// TwinCAT 3 PLC project WFServer
// ProgramVersion: 3.1.4026.14
// libraries:
//   Tc2_Standard, * (Beckhoff Automation GmbH)
//   Tc2_System, * (Beckhoff Automation GmbH)
//   Tc2_TcpIp, * (Beckhoff Automation GmbH)
//   Tc2_Utilities, * (Beckhoff Automation GmbH)
//   Tc3_Acsi, * (Beckhoff Automation GmbH)
//   Tc3_Ber, * (Beckhoff Automation GmbH)
//   Tc3_Collections, * (Beckhoff Automation GmbH)
//   Tc3_EventLogger, * (Beckhoff Automation GmbH)
//   Tc3_Gse, * (Beckhoff Automation GmbH)
//   Tc3_iec61850, * (Beckhoff Automation GmbH)
//   Tc3_iec61850_8_1, * (Beckhoff Automation GmbH)
//   Tc3_Mms, * (Beckhoff Automation GmbH)
//   Tc3_Rfc1006, * (Beckhoff Automation GmbH)
//   Tc3_Sockets, * (Beckhoff Automation GmbH)
//   Tc3_Tpkt, * (Beckhoff Automation GmbH)
//   Tc3_Ulosi, * (Beckhoff Automation GmbH)
// project tree:
//   / CommHandlerTask.TcTTO, DH_TCP_TX_TASK.TcTTO, IEC61850_TASK.TcTTO, UDP_RX_TASK.TcTTO, UDP_TX_TASK.TcTTO
//   DUTs/IEC61850/ E_DirectControlState.TcDUT, E_SboControlState.TcDUT
//   DUTs/IEC61850/User61850Enums/ E_ClrOp.TcDUT, E_CtlMd.TcDUT, E_TurCtl.TcDUT
//   DUTs/ S_TURBINECMD.TcDUT, S_TURBINEDATA.TcDUT
//   DUTs/TCP_UDP/ E_TCPConnectionState.TcDUT, E_UDPClientServerState.TcDUT, ST_TCPBinaryFrame.TcDUT, ST_TCPBinaryHeader.TcDUT, ST_UDPFrameEntry.TcDUT, TCP_DATA.TcDUT, UDP_DATA.TcDUT
//   GVLs/ CONSTANTS.TcGVL, TCP_GLOBALS.TcGVL, TcTelecontrol.TcGVL, UDP_GLOBALS.TcGVL
//   POUs/Common/ FB_LogFifo.TcPOU
//   POUs/COMM/ F_CreateTurbineCMD.TcPOU, F_InsertTurbineDataIEC61850.TcPOU, ParseTurbineData.TcPOU
//   POUs/ DH_TX_TCP_MAIN.TcPOU, P_IEC61850_MAIN.TcPOU, P_COMM_HANDLER.TcPOU, UDP_RX_MAIN.TcPOU, UDP_TX_MAIN.TcPOU
//   POUs/IEC61850Server/ FB_Control.TcPOU, FB_DirectControl.TcPOU, FB_DirectControlEnhanced.TcPOU, FB_SboControl.TcPOU, FB_SboControlEnhanced.TcPOU, FB_WTURBINEGse.TcPOU, FB_WTURBINEServerSession.TcPOU, FB_IEC61850.TcPOU, F_IEC61850ServerInit.TcPOU
//   POUs/IEC61850Server/User61850Enums/ FB_ClrOp.TcPOU, FB_CtlMd.TcPOU, FB_TurCtl.TcPOU
//   POUs/IEC61850Server/Util/ F_BuildAPTitle.TcPOU, F_BuildSelector.TcPOU, F_UdintToStringPadded.TcPOU
//   POUs/IEC61850Server/WTURBINE/ FB_IED_WTURBINE.TcPOU
//   POUs/IEC61850Server/WTURBINE/LD0/ FB_LD_WTURBINELD0.TcPOU
//   POUs/IEC61850Server/WTURBINE/LD0/LLN0/CDCs/ FB_DO_WTURBINE_LD0_LLN0_Beh.TcPOU, FB_DO_WTURBINE_LD0_LLN0_Health.TcPOU, FB_DO_WTURBINE_LD0_LLN0_Mod.TcPOU, FB_DO_WTURBINE_LD0_LLN0_NamPlt.TcPOU
//   POUs/IEC61850Server/WTURBINE/LD0/LLN0/ FB_LN_WTURBINE_LD0_LLN0.TcPOU
//   POUs/IEC61850Server/WTURBINE/LD0/LPHD1/CDCs/ FB_DO_WTURBINE_LD0_LPHD1_PhyHealth.TcPOU, FB_DO_WTURBINE_LD0_LPHD1_PhyNam.TcPOU, FB_DO_WTURBINE_LD0_LPHD1_Proxy.TcPOU
//   POUs/IEC61850Server/WTURBINE/LD0/LPHD1/ FB_LN_WTURBINE_LD0_LPHD1.TcPOU
//   POUs/IEC61850Server/WTURBINE/LD0/WALM1/CDCs/ FB_DO_WTURBINE_LD0_WALM1_Beh.TcPOU
//   POUs/IEC61850Server/WTURBINE/LD0/WALM1/ FB_LN_WTURBINE_LD0_WALM1.TcPOU
//   POUs/IEC61850Server/WTURBINE/LD0/WCNV1/CDCs/ FB_DO_WTURBINE_LD0_WCNV1_Beh.TcPOU, FB_DO_WTURBINE_LD0_WCNV1_Torq.TcPOU
//   POUs/IEC61850Server/WTURBINE/LD0/WCNV1/ FB_LN_WTURBINE_LD0_WCNV1.TcPOU
//   POUs/IEC61850Server/WTURBINE/LD0/WGEN1/CDCs/ FB_DO_WTURBINE_LD0_WGEN1_Beh.TcPOU, FB_DO_WTURBINE_LD0_WGEN1_RotSpd.TcPOU
//   POUs/IEC61850Server/WTURBINE/LD0/WGEN1/ FB_LN_WTURBINE_LD0_WGEN1.TcPOU
//   POUs/IEC61850Server/WTURBINE/LD0/WMET1/CDCs/ FB_DO_WTURBINE_LD0_WMET1_Beh.TcPOU, FB_DO_WTURBINE_LD0_WMET1_HorWdDir.TcPOU, FB_DO_WTURBINE_LD0_WMET1_HorWdSpd.TcPOU
//   POUs/IEC61850Server/WTURBINE/LD0/WMET1/ FB_LN_WTURBINE_LD0_WMET1.TcPOU
//   POUs/IEC61850Server/WTURBINE/LD0/WPPD1/CDCs/ FB_DO_WTURBINE_LD0_WPPD1_Beh.TcPOU, FB_DO_WTURBINE_LD0_WPPD1_ClrOp.TcPOU, FB_DO_WTURBINE_LD0_WPPD1_ClrOp_st.TcPOU, FB_DO_WTURBINE_LD0_WPPD1_DevOp.TcPOU, FB_DO_WTURBINE_LD0_WPPD1_DevOp_st.TcPOU, FB_DO_WTURBINE_LD0_WPPD1_DevSt.TcPOU, FB_DO_WTURBINE_LD0_WPPD1_DevSt_st.TcPOU
//   POUs/IEC61850Server/WTURBINE/LD0/WPPD1/DataSets/ FB_DS_TEMPLATE_LD1_WPPD1_ds01.TcPOU
//   POUs/IEC61850Server/WTURBINE/LD0/WPPD1/ FB_LN_WTURBINE_LD0_WPPD1.TcPOU
//   POUs/IEC61850Server/WTURBINE/LD0/WROT1/CDCs/ FB_DO_WTURBINE_LD0_WROT1_Beh.TcPOU, FB_DO_WTURBINE_LD0_WROT1_BlPthAngTgt.TcPOU, FB_DO_WTURBINE_LD0_WROT1_BlPthAngVal.TcPOU, FB_DO_WTURBINE_LD0_WROT1_RotSpd.TcPOU
//   POUs/IEC61850Server/WTURBINE/LD0/WROT1/ FB_LN_WTURBINE_LD0_WROT1.TcPOU
//   POUs/IEC61850Server/WTURBINE/LD0/WTUR1/CDCs/ FB_DO_WTURBINE_LD0_WTUR1_Beh.TcPOU, FB_DO_WTURBINE_LD0_WTUR1_DmdWSpt.TcPOU, FB_DO_WTURBINE_LD0_WTUR1_DmdWSpt_val.TcPOU, FB_DO_WTURBINE_LD0_WTUR1_TotWh.TcPOU, FB_DO_WTURBINE_LD0_WTUR1_TotWh_cntVal.TcPOU, FB_DO_WTURBINE_LD0_WTUR1_TurCtl.TcPOU, FB_DO_WTURBINE_LD0_WTUR1_TurCtl_st.TcPOU, FB_DO_WTURBINE_LD0_WTUR1_TurOp.TcPOU, FB_DO_WTURBINE_LD0_WTUR1_TurOp_st.TcPOU, FB_DO_WTURBINE_LD0_WTUR1_TurSt.TcPOU, FB_DO_WTURBINE_LD0_WTUR1_TurSt_st.TcPOU, FB_DO_WTURBINE_LD0_WTUR1_W.TcPOU
//   POUs/IEC61850Server/WTURBINE/LD0/WTUR1/ FB_LN_WTURBINE_LD0_WTUR1.TcPOU
//   POUs/IEC61850Server/WTURBINE/LD0/WYAW1/CDCs/ FB_DO_WTURBINE_LD0_WYAW1_Beh.TcPOU, FB_DO_WTURBINE_LD0_WYAW1_CabWup.TcPOU, FB_DO_WTURBINE_LD0_WYAW1_YwAng.TcPOU, FB_DO_WTURBINE_LD0_WYAW1_YwAngSpt.TcPOU, FB_DO_WTURBINE_LD0_WYAW1_YwAngSpt_val.TcPOU
//   POUs/IEC61850Server/WTURBINE/LD0/WYAW1/ FB_LN_WTURBINE_LD0_WYAW1.TcPOU
//   POUs/TCP/ FB_TCPClientConnection.TcPOU, FB_TCPClient.TcPOU, FB_TCPClientApplication.TcPOU
//   POUs/TCP/Util/ FB_TCPFrameFifo.TcPOU
//   POUs/UDP/ FB_UDPRxStateMachine.TcPOU, FB_UDPTxStateMachine.TcPOU
//   POUs/UDP/Util/ FB_UDPFrameFIFO.TcPOU
// real-time tasks:
//   TASK UDP_RX_TASK: cycle T#10ms, priority 15, ADS port 351
//   TASK CommHandlerTask: cycle T#10ms, priority 18, ADS port 353
//   TASK UDP_TX_TASK: cycle T#10ms, priority 2, ADS port 352
//   TASK IEC61850_TASK: cycle T#10ms, priority 1, ADS port 350
//   TASK DH_TCP_TX_TASK: cycle T#10ms, priority 3, ADS port 354
// I/O:
//   DEVICE GSE (RT-Ethernet Adapter) (disabled)

CONFIGURATION WFServer
    RESOURCE PLC ON TwinCAT3
        TASK CommHandlerTask(INTERVAL := T#10ms, PRIORITY := 18);
        TASK DH_TCP_TX_TASK(INTERVAL := T#10ms, PRIORITY := 3);
        TASK IEC61850_TASK(INTERVAL := T#10ms, PRIORITY := 1);
        TASK UDP_RX_TASK(INTERVAL := T#10ms, PRIORITY := 15);
        TASK UDP_TX_TASK(INTERVAL := T#10ms, PRIORITY := 2);
        PROGRAM P_COMM_HANDLER WITH CommHandlerTask : P_COMM_HANDLER;
        PROGRAM DH_TX_TCP_MAIN WITH DH_TCP_TX_TASK : DH_TX_TCP_MAIN;
        PROGRAM P_IEC61850_MAIN WITH IEC61850_TASK : P_IEC61850_MAIN;
        PROGRAM UDP_RX_MAIN WITH UDP_RX_TASK : UDP_RX_MAIN;
        PROGRAM UDP_TX_MAIN WITH UDP_TX_TASK : UDP_TX_MAIN;
    END_RESOURCE
END_CONFIGURATION

// ---- DUTs/IEC61850/E_DirectControlState.TcDUT
{attribute 'qualified_only'}
{attribute 'strict'}
TYPE E_DirectControlState : 
(
	Ready := 0,
	WaitForActivationTime := 1,
	PerformTest := 2,
	WaitForExecution := 3,
	Operate := 4,
	WaitForChange := 5,
	MirrorBlockedCommand := 6
) ;
END_TYPE

// ---- DUTs/IEC61850/E_SboControlState.TcDUT
{attribute 'qualified_only'}
{attribute 'strict'}
TYPE E_SboControlState : 
(
	Unselected := 0,
	Select_PerformTest := 1,
	WaitForSelection := 2,
	Ready := 3,
	WaitForActivationTime := 4,
	PerformTest := 5,
	WaitForExecution := 6,
	MirrorBlockedCommand := 7,
	Operate := 8,
	WaitForChange := 9,
	EndSelection := 10
) ;
END_TYPE

// ---- DUTs/IEC61850/User61850Enums/E_ClrOp.TcDUT
{attribute 'qualified_only'}
{attribute 'strict'}
TYPE E_ClrOp : 
(
	e_0 := 0, (*None*)
	e_1 := 1 (*Clear*)
) SINT;
END_TYPE

// ---- DUTs/IEC61850/User61850Enums/E_CtlMd.TcDUT
{attribute 'qualified_only'}
{attribute 'strict'}
TYPE E_CtlMd : 
(
	e_1 := 1, (*local*)
	e_2 := 2, (*remote*)
	e_3 := 3, (*auto*)
	e_4 := 4 (*test*)
) SINT;
END_TYPE

// ---- DUTs/IEC61850/User61850Enums/E_TurCtl.TcDUT
{attribute 'qualified_only'}
{attribute 'strict'}
TYPE E_TurCtl : 
(
	e_1 := 1, (*ROSCO*)
	e_2 := 2 (*Lio*)
) SINT;
END_TYPE

// ---- DUTs/S_TURBINECMD.TcDUT
(* Holds the command for all turbines *)
{attribute 'pack_mode' := '1'}
TYPE S_TURBINECMD :
STRUCT
	bEnable 		: ARRAY[1..c_nNumTurbines] OF BOOL;
	bEmergencyStop	: ARRAY[1..c_nNumTurbines] OF BOOL;
	eCtrlMode		: ARRAY[1..c_nNumTurbines] OF SINT;		// 1 Byte
	fWSpt			: ARRAY[1..c_nNumTurbines] OF REAL;
	fYawSpt			: ARRAY[1..c_nNumTurbines] OF REAL;
END_STRUCT
END_TYPE

// ---- DUTs/S_TURBINEDATA.TcDUT
{attribute 'pack_mode' := '1'}
TYPE S_TURBINEDATA :
STRUCT
	WindSpeed			: REAL;
	WindDirection		: REAL;
	PowerGen			: REAL;
	YawAng				: REAL;
	RotorSpeed			: REAL;
	PitchAngle			: REAL;
	PitchAngleSpt		: REAL;
	GenTorque			: REAL;
END_STRUCT
END_TYPE

// ---- DUTs/TCP_UDP/E_TCPConnectionState.TcDUT
TYPE E_TCPConnectionState :
(
	eTCP_STATE_IDLE,
	eTCP_STATE_CONNECT_START,
	eTCP_STATE_CONNECT_WAIT,
	eTCP_STATE_DATAEXCHANGE,
	eTCP_STATE_CLOSE_START,
	eTCP_STATE_CLOSE_WAIT,
	eTCP_STATE_ERROR
);
END_TYPE

// ---- DUTs/TCP_UDP/E_UDPClientServerState.TcDUT
TYPE E_UDPClientServerState :
(
	eUDP_STATE_IDLE		:= 0,
	eUDP_STATE_CREATE_START,
	eUDP_STATE_CREATE_WAIT,
	eUDP_STATE_SEND_START,
	eUDP_STATE_SEND_WAIT,
	eUDP_STATE_RECEIVE_START,
	eUDP_STATE_RECEIVE_WAIT,
	eUDP_STATE_CLOSE_START,
	eUDP_STATE_CLOSE_WAIT,
	eUDP_STATE_ERROR
);
END_TYPE

// ---- DUTs/TCP_UDP/ST_TCPBinaryFrame.TcDUT
(* Simple binary TCP/IP frame (8 byte aligned) *)
TYPE ST_TCPBinaryFrame :
STRUCT
	head	: ST_TCPBinaryHeader;(* Frame header (16 byte) *)
	data 	: TCP_DATA;(* User data (?? byte) *)

	(* Total frame size = 16+?? byte *)
END_STRUCT
END_TYPE

// ---- DUTs/TCP_UDP/ST_TCPBinaryHeader.TcDUT
(* Simple binary TCP/IP frame header (8 byte aligned) *)
TYPE ST_TCPBinaryHeader :
STRUCT
	dwStart		: DWORD	:= 16#BECF1234;	(* Start bytes *)
	cbLength	: UDINT(0..cTCP_BUFFER_SIZE) := 0;(* Max. length of attached binary data *)
	nS			: UDINT := 0;(* Send counter *)
	nR			: UDINT	:= 0;(* Receive counter *)
	
	(* Total header data size = 16 byte *)
END_STRUCT
END_TYPE

// ---- DUTs/TCP_UDP/ST_UDPFrameEntry.TcDUT
TYPE ST_UDPFrameEntry :
STRUCT
	stRemoteAddr 	: ST_SockAddr;	(* Remote address. String containing an (Ipv4) Internet Protocol dotted address and port number. *)
	sMessage		: UDP_DATA;	(* UDP packet data *)
END_STRUCT
END_TYPE

// ---- DUTs/TCP_UDP/TCP_DATA.TcDUT
// TYPE TCP_DATA : ARRAY[1..cTCP_FrameSize] OF BYTE; END_TYPE
TYPE TCP_DATA :
STRUCT
	nID				: UDINT;
	nUnixTime		: ULINT;
	YwAng			: REAL;
	YwAngSpt		: REAL;
	W				: REAL;
	WSpt			: REAL;
	HorWdSpd		: REAL;
	HorWdDir		: REAL;
	RotSpd			: REAL;
	PitchAngle		: REAL;
	PitchAngleSpt	: REAL;
// 	GenTorque		: REAL;
END_STRUCT
END_TYPE

// ---- DUTs/TCP_UDP/UDP_DATA.TcDUT
TYPE UDP_DATA : ARRAY[1..SIZEOF(S_TURBINECMD)*c_nNumTurbines] OF BYTE; END_TYPE

// ---- GVLs/CONSTANTS.TcGVL
VAR_GLOBAL CONSTANT
	c_nNumTurbines	: UDINT := 9;
	
	(* IEC 61850 Server Definitions *)
	c_aIpAddr 		: STRING := '172.19.3.190';
	c_aMMSPortBase 	: UDINT := 102;
	c_aAP_invIDBase : INT := 0;
	c_nNumSessions	: UINT := 1;
	
	(* UDP Connection Constants *)
	sSrvNetId			: T_AmsNetID 	:= '';(* TwinCAT TCP/IP server network address. Default: empty string. *)
	sLocalHost			: T_IPv4Addr 	:= '172.19.3.190';(* Local address: String containing an (Ipv4) Internet Protocol dotted address. *)
	nLocalTxPort		: UDINT			:= 11000;	(* UDP port used for transmission *)
	nLocalRxPort		: UDINT			:= 11001;	(* UDP port used for receiving *)
	sRemoteHost			: T_IPv4Addr 	:= '172.19.3.43';(* Remote address: String containing an (Ipv4) Internet Protocol dotted address. *)
	nRemoteTxPort		: UDINT 		:= 11000; (* Remote address: IP Tx port number. *)
	nRemoteRxPort		: UDINT			:= 10000; (* Remote address: IP Rx port number. *)
	
	UDP_RX_BUFFER_SIZE 	: UDINT := c_nNumTurbines * 1024; 	// Size of the UDP RX FIFO Buffer in Bytes
	UDP_TX_BUFFER_SIZE 	: UDINT := 1024; 	// Size of the UDP TX FIFO Buffer in Bytes
	
	UDP_ERR_TX_FIFO_OF	: UDINT := 16#8103;
	UDP_ERR_RX_FIFO_OF	: UDINT := 16#8104;
END_VAR

// ---- GVLs/TCP_GLOBALS.TcGVL
VAR_GLOBAL CONSTANT
	cTCP_BUFFER_SIZE						: UDINT := 1000;
	cTCP_FrameSize							: UDINT := 256;

	cTCP_SEND_CYCLE_TIME					: TIME := T#1S;
	cTCP_RECEIVE_POLLING_TIME		 		: TIME := T#100MS;
	cTCP_RECEIVE_TIMEOUT					: TIME := T#50S;

	(* Some project specific error codes *)
	cTCP_ERROR_RECEIVE_TIMEOUT				: UDINT := 16#8101;(* Receive timeout error *)
	cTCP_ERROR_SENDFIFO_OVERFLOW			: UDINT := 16#8102;(* Send fifo overflow *)
	cTCP_ERROR_RECFIFO_OVERFLOW				: UDINT := 16#8103;(* Receive fifo overflow *)
	cTCP_ERROR_INVALID_FRAME_FORMAT		: UDINT := 16#8104;(* Invalid frame format/data *)
END_VAR

// ---- GVLs/TcTelecontrol.TcGVL
VAR_GLOBAL
	ipCreator: I_AcsiCodeCreatorClass := GVL_AcsiVars.Creator.SetCodeRev(codeRev:=7).SetGuiVer(major:=3, minor:=98, build:=20, revision:=0);
	
	(* IEC61850 Data Models for Turbine *)
	fbWTURBINE: ARRAY[1..c_nNumTurbines] OF FB_IED_WTURBINE;
	
	(* IEC61850 Server Objects, one for each turbine *)
	fbServer : ARRAY[1..c_nNumTurbines] OF FB_iec61850ServerClass;
	
	(* IEC61850 Server Sessions, one or multiple for each server object *)
	fbSession: ARRAY[1..c_nNumTurbines, 1..c_nNumSessions] OF FB_WTURBINEServerSession;
	
// 	{warning 'Please configure your server IP-address in the initialization code of the server function block below:'}
	(* Server container *)
// 	fbWTURBINEServer: FB_iec61850ServerClass := (ipIED:=fbWTURBINE, settings:=(bEnable:=TRUE, sLocalHost:='192.168.1.100', nCalled_AP_InvID:=0, nCalling_AP_InvID:=0, nCalled_AE_InvID:=0, nCalling_AE_InvID:=0));
	
	(* Server connections *)
// 	fbWTURBINEServerSession1: FB_WTURBINEServerSession := (fbConnection:=(ipServer:=fbWTURBINEServer, settings:=(bEnable:=TRUE)));
	(*
	fbWTURBINEServerSession2: FB_WTURBINEServerSession := (fbConnection:=(ipServer:=fbWTURBINEServer, settings:=(bEnable:=TRUE)));
	...
	fbWTURBINEServerSessionN: FB_WTURBINEServerSession := (fbConnection:=(ipServer:=fbWTURBINEServer, settings:=(bEnable:=TRUE)));
	*)
	
	
// 	fbWTURBINEGse: FB_WTURBINEGse := (fbAdapter:=(ipIED:=fbWTURBINE, settings:=(sMulticastAddr:='01-0C-CD-01-00-00', eDispatchMode:=E_GseDispatchMode.NonPromiscuous)));
	
	
END_VAR

// ---- GVLs/UDP_GLOBALS.TcGVL
VAR_GLOBAL
	(* Global TX and RX buffers, together with their respective critical section handlers*)
// 	fbUDP_RX_CS			: FB_IecCriticalSection;
	fbRxFIFO			: FB_UDPFrameFIFO;
	
// 	fbUDP_TX_CS			: FB_IecCriticalSection;
	fbTxFIFO			: FB_UDPFrameFIFO;
END_VAR

// ---- POUs/P_COMM_HANDLER.TcPOU
PROGRAM P_COMM_HANDLER
VAR
	i					: UDINT;
	nAddr				: ULINT;
	stReceivedFrom		: ST_UDPFrameEntry;
	sLoggedMessage		: UDP_DATA;
	dVal_1				: LREAL;
	dVal_2				: LREAL;	
	sTurbineData		: S_TURBINEDATA;
	iTemp				: ULINT;
	
	sTxTimer			: TON;
	bSend				: BOOL := FALSE;
	cTxTimerPeriod		: TIME := T#500MS;
	sTurbineCmd			: S_TURBINECMD;
	stSendTo			: ST_UDPFrameEntry;;
END_VAR


(* First we pop from the UDP RX buffer, and process the received data accordingly *)
REPEAT
	fbRxFIFO.RemoveHead( );
	IF fbRxFIFO.bOk THEN

		(* TODO:: Implement received frame handler *)
		stReceivedFrom := fbRxFIFO.stGet;
		IF stReceivedFrom.stRemoteAddr.sAddr = sRemoteHost AND stReceivedFrom.stRemoteAddr.nPort = nRemoteTxPort THEN
// 			sLoggedMessage := stReceivedFrom.sMessage;
			nAddr := 0;
			FOR i := 1 TO c_nNumTurbines DO
				sTurbineData := ParseTurbineData(ADR(stReceivedFrom.sMessage) + nAddr);
				F_InsertTurbineDataIEC61850(nID := i, sTurbineData := sTurbineData);
				nAddr := nAddr + SIZEOF(S_TURBINEDATA);
			END_FOR
		END_IF
// 		MEMCPY(ADR(dVal_1), ADR(sLoggedMessage), SIZEOF(dVal_1));
// 		MEMCPY(ADR(dVal_2), ADR(sLoggedMessage) + SIZEOF(dVal_1), SIZEOF(dVal_2));
// 			ADSLOGSTR( ADSLOG_MSGTYPE_HINT OR ADSLOG_MSGTYPE_LOG OR ADSLOG_MSGTYPE_MSGBOX, '%s', stReceivedFrom.sMessage );
		
	END_IF
UNTIL NOT fbRxFIFO.bOk
END_REPEAT


(* Second, we take the turbine setpoints and transmit to the turbine *)
bSend := sTxTimer.Q;
sTxTimer(IN := NOT sTxTimer.Q, PT := cTxTimerPeriod);

IF bSend THEN
	sTurbineCmd := F_CreateTurbineCMD();
	fbTXFIFO.AddTail( );
	iTemp :=  SIZEOF(sTurbineCmd);
	MEMCPY(ADR(stSendTo.sMessage), ADR(sTurbineCmd), SIZEOF(sTurbineCmd));
	stSendTo.stRemoteAddr.sAddr := sRemoteHost;	(* Remote host IP address *)
	stSendTo.stRemoteAddr.nPort := nRemoteRxPort;	(* Remote host port number *)
	fbTxFIFO.AddTail( stPut := stSendTo );
END_IF

END_PROGRAM

// ---- POUs/COMM/ParseTurbineData.TcPOU
FUNCTION ParseTurbineData
VAR_INPUT
	sMessage		: POINTER TO BYTE;
END_VAR
VAR_OUTPUT
	sTurbineData	: S_TURBINEDATA;
// 	bOk				: BOOL;
END_VAR
VAR
	i				: UDINT;
	nAddr			: ULINT;
END_VAR

// bOk := FALSE;
MEMCPY(ADR(sTurbineData), sMessage, SIZEOF(sTurbineData));
// nAddr := 0;
// MEMCPY(ADR(sTurbineData.WindSpeed) + nAddr, sMessage + nAddr, SIZEOF(sTurbineData.WindSpeed));
// nAddr := nAddr + SIZEOF(sTurbineData.WindSpeed);
// 
// MEMCPY(ADR(sTurbineData.WindDirection), sMessage + nAddr, SIZEOF(sTurbineData.WindDirection));
// nAddr := nAddr + SIZEOF(sTurbineData.WindDirection);
// 
// MEMCPY(ADR(sTurbineData.PowerGen), sMessage + nAddr, SIZEOF(sTurbineData.PowerGen));
// nAddr := nAddr + SIZEOF(sTurbineData.PowerGen);
// 
// MEMCPY(ADR(sTurbineData.YawAng), sMessage + nAddr, SIZEOF(sTurbineData.YawAng));
// nAddr := nAddr + SIZEOF(sTurbineData.YawAng);
// 
// MEMCPY(ADR(sTurbineData.RotorSpeed), sMessage + nAddr, SIZEOF(sTurbineData.RotorSpeed));
// nAddr := nAddr + SIZEOF(sTurbineData.RotorSpeed);
// 
// MEMCPY(ADR(sTurbineData.PitchAngle), sMessage + nAddr, SIZEOF(sTurbineData.PitchAngle));
// nAddr := nAddr + SIZEOF(sTurbineData.PitchAngle);
// 
// MEMCPY(ADR(sTurbineData.PitchAngleSpt), sMessage + nAddr, SIZEOF(sTurbineData.PitchAngleSpt));
// nAddr := nAddr + SIZEOF(sTurbineData.PitchAngleSpt);
// 
// MEMCPY(ADR(sTurbineData.GenTorque), sMessage + nAddr, SIZEOF(sTurbineData.GenTorque));
// nAddr := nAddr + SIZEOF(sTurbineData.GenTorque);

// bOk := TRUE;

END_FUNCTION

// ---- POUs/COMM/F_InsertTurbineDataIEC61850.TcPOU
FUNCTION F_InsertTurbineDataIEC61850
VAR_INPUT
	nID				: UDINT;
	sTurbineData	: S_TURBINEDATA;
END_VAR
VAR_OUTPUT
END_VAR
VAR
END_VAR

IF nID >= 1 OR nID <= c_nNumTurbines THEN
	fbWTURBINE[nID].WTURBINELD0.WMET1.HorWdSpd.mag.fValue := sTurbineData.WindSpeed;
	fbWTURBINE[nID].WTURBINELD0.WMET1.HorWdDir.mag.fValue := sTurbineData.WindDirection;
	fbWTURBINE[nID].WTURBINELD0.WTUR1.W.mag.fValue := sTurbineData.PowerGen;
	fbWTURBINE[nID].WTURBINELD0.WYAW1.YwAng.mag.fValue := sTurbineData.YawAng;
	fbWTURBINE[nID].WTURBINELD0.WROT1.RotSpd.mag.fValue := sTurbineData.RotorSpeed;
	fbWTURBINE[nID].WTURBINELD0.WROT1.BlPthAngVal.mag.fValue := sTurbineData.PitchAngle;
	fbWTURBINE[nID].WTURBINELD0.WROT1.BlPthAngTgt.mag.fValue := sTurbineData.PitchAngleSpt;
 	fbWTURBINE[nID].WTURBINELD0.WCNV1.Torq.mag.fValue := sTurbineData.GenTorque;
END_IF

END_FUNCTION

// ---- POUs/COMM/F_CreateTurbineCMD.TcPOU
FUNCTION F_CreateTurbineCMD
VAR_INPUT
// 	nID				: UDINT;
END_VAR
VAR_OUTPUT
	sTurbineCmd		: S_TURBINECMD;
END_VAR
VAR
	temp: SINT;
	nID: UDINT;
END_VAR


FOR nID := 1 TO c_nNumTurbines DO
	temp := fbWTURBINE[nID].WTURBINELD0.WTUR1.TurOp.st_.stVal.iAny;
	sTurbineCmd.bEnable[nID] :=  SINT_TO_BOOL(temp);
	sTurbineCmd.bEmergencyStop[nID] := FALSE;
	sTurbineCmd.eCtrlMode[nID] := fbWTURBINE[nID].WTURBINELD0.WTUR1.TurCtl.st_.stVal.iAny;
	sTurbineCmd.fWSpt[nID] 	:= fbWTURBINE[nID].WTURBINELD0.WTUR1.DmdWSpt.val.mxVal.fValue;
	sTurbineCmd.fYawSpt[nID] := fbWTURBINE[nID].WTURBINELD0.WYAW1.YwAngSpt.val.mxVal.fValue;
END_FOR

END_FUNCTION

// ---- POUs/DH_TX_TCP_MAIN.TcPOU
PROGRAM DH_TX_TCP_MAIN
VAR
	sSrvNetID 	: T_AmsNetID := '';(* TwinCAT TCP/IP server network address *)
	bEnable 	: BOOL := TRUE;(* TRUE => Enable client data exchange, FALSE => Disable *)	
	
	bLog		: BOOL := TRUE;(* TRUE => Enable message/error log, FALSE => Disable*)
	
	fbClient : FB_TCPClient := ( sRemoteHost:= '172.19.3.214',(* IP address of remote server! *)
								nRemotePort:= 9003,(* Port number of remote server! *)
								sPrefix := 'CLIENT1::' );(* TCP/IP client (connection) instance *)
								
	fbCloseAll		: FB_SocketCloseAll;
	bInitialize		: BOOL := TRUE;
END_VAR

IF fbCloseAll.bBusy OR fbCloseAll.bError THEN
	RETURN;
END_IF
bInitialize := FALSE;

fbClient( sSrvNetID := sSrvNetID, bEnable := bEnable, bLog := bLog );

END_PROGRAM

// ---- POUs/TCP/FB_TCPClient.TcPOU
FUNCTION_BLOCK FB_TCPClient
VAR_INPUT
	sSrvNetID	: T_AmsNetID	:= '';(* TwinCAT TCP/IP server network address *)
	sRemoteHost	: T_IPv4Addr 	:= '127.0.0.1';(* Server IP network address *)
	nRemotePort	: UDINT 		:= 200;(* Server port number *)
	bEnable		: BOOL 			:= FALSE;(* TRUE => enable client data exchange, FALSE => disable *)
	bLog		: BOOL 			:= FALSE;(* TRUE => Enable log message output, FALSE => Disable *)
	sPrefix		: STRING 		:= 'CLIENT::';(* Log message description string (allows the identification of log message source) *)
END_VAR
VAR_OUTPUT
	eState		: E_SocketConnectionState := eSOCKET_DISCONNECTED;(* TCP/IP connection state *)
END_VAR
VAR
	fbApplication 	: FB_TCPClientApplication;(* Client application control function block *)
	fbConnection	: FB_TCPClientConnection;(* Client data exchange control function block *)
	fbTx 			: FB_TCPFrameFifo;(* Tx fifo *)
	fbRx 			: FB_TCPFrameFifo;(* Rx fifo *)
	fbLog			: FB_LogFifo;(* Log/debug/error fifo *)
END_VAR

(*-------------------------- Trigger data exchange -----------------------------------------------*)
fbConnection( 	sSrvNetID := sSrvNetID, fbRx := fbRx, fbTx := fbTx, fbLog := fbLog, 
				bEnable := bEnable, sRemoteHost := sRemoteHost, nRemotePort := nRemotePort,  
				bLog := bLog, sPrefix := sPrefix, eState=>eState );
	
IF fbConnection.eState = eSOCKET_CONNECTED THEN(* Connection established *)
	fbApplication( fbTx := fbTx, fbRx := fbRx, fbLog := fbLog );
END_IF

END_FUNCTION_BLOCK

// ---- POUs/TCP/FB_TCPClientApplication.TcPOU
FUNCTION_BLOCK FB_TCPClientApplication
VAR_IN_OUT
	fbTx 		: FB_TCPFrameFifo;(* TX fifo *)
	fbRx 		: FB_TCPFrameFifo;(* RX fifo *)
	fbLog		: FB_LogFifo;(* Log message fifo *)
END_VAR
VAR
	stToServer	: TCP_DATA;
	stFromServer: TCP_DATA;
	sLogMessage	: T_MaxString := '';
	nCounter	: UDINT;
	fbSndTimer	: TON;
	i: UDINT;
	fbFormat   : FB_FormatString;
	sFormatted : T_MaxString;
	
	
	fbTime   : FB_LocalSystemTime := ( bEnable := TRUE, dwCycle := 1 );
	sTime 	: T_MaxString;
 	nDataLen     : INT;
    nUnixTime    : LINT;
END_VAR

(*------------------- Send cyclic message strings ------------------------------------*)
(* TODO: Make this 'application/task' agnostic. *)
(* For now, it always sends logging data to the historian *)
fbSndTimer( IN := TRUE, PT := cTCP_SEND_CYCLE_TIME );
IF fbSndTimer.Q THEN(* Send string to server *)
	fbSndTimer( IN := FALSE );

// 	nCounter := nCounter  + 1;
// 	stToServer := MAXSTRING_TO_BYTEARR(CONCAT( 'Client message: ', UDINT_TO_STRING(nCounter) ));
//  
// 	fbTx.AddTail( stPut := stToServer );(* Put string to the tx fifo *)
// 	IF NOT fbTx.bOk THEN(* TX fifo overflow => log error *)
// 		fbLog.Error( sMessage := 'FB_FrameFifo(sender)\0', nErrID := cTCP_ERROR_SENDFIFO_OVERFLOW );
// 	END_IF
	
	fbTime();
	sTime := SYSTEMTIME_TO_STRING(fbTime.systemTime);
	FOR i := 1 TO c_nNumTurbines DO
		
		stToServer.nID := i;
		stToServer.nUnixTime := (F_GetSystemTime() - 116444736000000000) / 10000000;
		stToServer.YwAng := fbWTURBINE[i].WTURBINELD0.WYAW1.YwAng.mag.fValue;
		stToServer.YwAngSpt := fbWTURBINE[i].WTURBINELD0.WYAW1.YwAngSpt.val.mxVal.fValue;
		stToServer.W := fbWTURBINE[i].WTURBINELD0.WTUR1.W.mag.fValue;
		stToServer.WSpt := fbWTURBINE[i].WTURBINELD0.WTUR1.DmdWSpt.val.mxVal.fValue;
		stToServer.HorWdSpd := fbWTURBINE[i].WTURBINELD0.WMET1.HorWdSpd.mag.fValue;
		stToServer.HorWdDir := fbWTURBINE[i].WTURBINELD0.WMET1.HorWdDir.mag.fValue;
		stToServer.RotSpd := fbWTURBINE[i].WTURBINELD0.WROT1.RotSpd.mag.fValue;
		stToServer.PitchAngle := fbWTURBINE[i].WTURBINELD0.WROT1.BlPthAngVal.mag.fValue;
		stToServer.PitchAngleSpt := fbWTURBINE[i].WTURBINELD0.WROT1.BlPthAngTgt.mag.fValue;
// 		stToServer.GenTorque := fbWTURBINE[i].WTURBINELD0.WROT1.
		
		
		
		
		fbTx.AddTail( stPut := stToServer );(* Put string to the tx fifo *)
		IF NOT fbTx.bOk THEN(* TX fifo overflow => log error *)
			fbLog.Error( sMessage := 'FB_FrameFifo(sender)\0', nErrID := cTCP_ERROR_SENDFIFO_OVERFLOW );
		END_IF
	END_FOR

END_IF

END_FUNCTION_BLOCK

// ---- POUs/TCP/Util/FB_TCPFrameFifo.TcPOU
(* Tx/Rx (string data) fifo control function block *)
FUNCTION_BLOCK FB_TCPFrameFifo
VAR_INPUT
	bLog		: BOOL		:= FALSE;(* TRUE => Enable log message output, FALSE => Disable *)
	sPrefix		: STRING	:= 'Unknown::';(* Log message description string (allows the identification of log message source) *)
	stPut		: TCP_DATA;(* Frame to add (write) to the fifo *)
END_VAR
VAR_OUTPUT
	bOk			: BOOL; 	(* TRUE = New entry added or removed succesfully, FALSE = Fifo overflow or fifo empty *)
	stGet		: TCP_DATA;(* Frame removed (read) from fifo *)
	nCount		: UDINT		:= 0;(* Number of fifo entries *)
	cbFree		: UDINT 	:= 0;(* Free buffer space *)
END_VAR
VAR
	fbBuffer 	: FB_MemRingBuffer;(* Basic (lower level) buffer control function block *)
	buffer		: ARRAY[-3..cTCP_BUFFER_SIZE] OF BYTE;(* Internal buffer memory *)
END_VAR

;

ACTION AddTail:
(* Adds new fifo entry *)
fbBuffer.A_AddTail( pBuffer:= ADR(buffer), cbBuffer:= SIZEOF(buffer),
					pWrite := ADR( stPut ), cbWrite := SIZEOF( stPut ), 
					bOk=>bOk, nCount=>nCount );
IF bOk THEN
	cbFree := cTCP_BUFFER_SIZE - fbBuffer.cbSize;(* Calculate the free buffer space *)
// 	IF bLog THEN(* Log message *)
// 		F_ADSLOGHEXDATA( CONCAT( sPrefix, '<=' ), ADR( stPut ), SIZEOF( stPut ) );
// 	END_IF
END_IF
END_ACTION

ACTION Clear:
(* Resets fifo = clears all data *)
MEMSET( ADR( stGet ), 0, SIZEOF( stGet ) );
fbBuffer.A_Reset( pBuffer:= ADR(buffer), cbBuffer:= SIZEOF(buffer),
					pWrite := ADR( stPut ), cbWrite := SIZEOF( stPut ), 
					pRead := ADR( stGet ), cbRead := SIZEOF( stPut ),
					bOk=>bOk, nCount=>nCount );
cbFree := cTCP_BUFFER_SIZE;(* Free buffer size *)
END_ACTION

ACTION RemoveHead:
(* Removes oldest fifo entry *)
MEMSET( ADR( stGet ), 0, SIZEOF( stGet ) );
fbBuffer.A_RemoveHead( pBuffer:= ADR(buffer), cbBuffer:= SIZEOF(buffer),
						pRead := ADR( stGet ), cbRead := SIZEOF( stGet ),
						bOk=>bOk, nCount=>nCount );
IF bOk THEN
	cbFree := cTCP_BUFFER_SIZE - fbBuffer.cbSize;(* Calculate the free buffer space *)
END_IF
END_ACTION

END_FUNCTION_BLOCK

// ---- POUs/Common/FB_LogFifo.TcPOU
(* Log/debug/error message fifo *)
FUNCTION_BLOCK FB_LogFifo
VAR_INPUT
	bLog		: BOOL 		:= FALSE;(* TRUE => Enable log message output, FALSE => Disable *)
	sPrefix		: STRING 	:= 'Unknown::';(* Log message description string (allows the identification of log message source) *)
	
	sMessage	: STRING 	:= '';(* String message to add (write) to the fifo *)
	nErrID		: UDINT 	:= 0;(* Error code to add (write) to the fifo *)
	hSocket		: T_HSOCKET;(* Socket connection handle *)
END_VAR
VAR_OUTPUT
	bOk			: BOOL;(* TRUE = New entry added or removed succesfully, FALSE = Fifo overflow or fifo empty *)
	sGet		: T_MaxString := '';(* String entry removed (read) from fifo *)
	nCount		: UDINT := 0;(* Number of fifo entries *)
END_VAR
VAR
	fbBuffer 	: FB_StringRingBuffer;(* Basic (lower level) string buffer control function block *)
	buffer		: ARRAY[0..cTCP_BUFFER_SIZE] OF BYTE;(* Internal buffer memory *)
	sSource		: T_MaxString;	
	sPut		: T_MaxString;
END_VAR

;

ACTION Clear:
(* Clears all fifo entries *)
fbBuffer.A_Reset( 	pBuffer := ADR( buffer ), cbBuffer := SIZEOF( buffer ), 
					bOk=>bOk, nCount=>nCount, getValue=>sGet );
END_ACTION

ACTION Error:
(* Adds new fifo entry *)
IF nErrID = 0 THEN
	sSource := '::Error: 0x';
ELSIF ( nErrID AND 16#80000000) = 16#80000000 THEN
	IF nErrID = 16#80072746 THEN
		sSource := '::Win32 error (the connection is reset by remote side): 0x';
	ELSE
		sSource := '::Win32 error: 0x';
	END_IF
ELSIF (nErrID AND 16#00008100) = 16#00008100 THEN
	CASE nErrID OF
		cTCP_ERROR_RECEIVE_TIMEOUT:
			sSource := '::PLC sample project receive timeout error: 0x';
		cTCP_ERROR_SENDFIFO_OVERFLOW:
			sSource := '::PLC sample project send fifo overflow error: 0x';
		cTCP_ERROR_RECFIFO_OVERFLOW:
			sSource := '::PLC sample project receive fifo overflow error: 0x';
	ELSE
		sSource := '::Other PLC sample project error: 0x';
	END_CASE
ELSIF (nErrID AND 16#00008000) = 16#00008000 THEN
	sSource := '::Internal TCP/IP Connection Server error: 0x';
ELSE
	sSource := '::TwinCAT System error: 0x';
END_IF

sPut := CONCAT( CONCAT( CONCAT( sPrefix, sMessage ), sSource ), DWORD_TO_HEXSTR( nErrID AND 16#FFFF, 0, FALSE ) ); 

fbBuffer.A_AddTail( pBuffer:= ADR(buffer), cbBuffer:= SIZEOF(buffer),
					putValue:= sPut, bOk=>bOk, nCount=>nCount );
IF bOk THEN
	IF bLog THEN(* Log error message *)
		ADSLOGSTR( ADSLOG_MSGTYPE_ERROR OR ADSLOG_MSGTYPE_LOG, '%s', sPut );	
	END_IF
END_IF
END_ACTION

ACTION Message:
(* Adds new fifo entry *)
sPut := CONCAT( CONCAT( sPrefix, sMessage ), CONCAT( '::', HSOCKET_TO_STRING(hSocket) ) );
fbBuffer.A_AddTail( pBuffer:= ADR(buffer), cbBuffer:= SIZEOF(buffer),
					putValue:= sPut, bOk=>bOk, nCount=>nCount );
IF bOk THEN
	IF bLog THEN(* Log information message *)
		ADSLOGSTR( ADSLOG_MSGTYPE_HINT OR ADSLOG_MSGTYPE_LOG, '%s', sPut );	
	END_IF
END_IF
END_ACTION

ACTION Remove:
(* Removes oldest fifo entry *)
IF nCount = 0 THEN
	sGet := '';
	bOk := FALSE;
	RETURN;
END_IF

fbBuffer.A_RemoveHead( pBuffer:= ADR(buffer), cbBuffer:= SIZEOF(buffer),
						getValue=>sGet, bOk=>bOk, nCount=>nCount );
END_ACTION

END_FUNCTION_BLOCK

// ---- POUs/TCP/FB_TCPClientConnection.TcPOU
(* 	This function block implements simple TCP/IP client protocol. *)
FUNCTION_BLOCK FB_TCPClientConnection
VAR_IN_OUT
	fbTx 		: FB_TCPFrameFifo;(* TX fifo *)
	fbRx 		: FB_TCPFrameFifo;(* RX fifo *)
	fbLog		: FB_LogFifo;(* Log message fifo *)
END_VAR
VAR_INPUT
	sSrvNetID	: T_AmsNetID	:= '';(* TwinCAT TCP/IP server network address *)
	sRemoteHost	: T_IPv4Addr 	:= '127.0.0.1';(* IP address of remote server *)
	nRemotePort	: UDINT			:= 200;(* Remote server port *)
	bEnable		: BOOL			:= FALSE;(* TRUE => Enable/connect, FALSE => Disable/disconnect *)
	tReconnect	: TIME 			:= T#5S;(* Try to reconnect after this time *)
	bLog		: BOOL 			:= FALSE; (* TRUE => Enable debug output, FALSE => Disable debug output *)
	sPrefix		: STRING 		:= 'CLIENT::';(* Log message description string (allows the identification of log message source) *)
END_VAR
VAR_OUTPUT
	eState		: E_SocketConnectionState := eSOCKET_DISCONNECTED;(* TCP/IP connection state *)
END_VAR
VAR
	fbConnect 	: FB_ClientServerConnection;(* Create/release TCP/IP connection *)
	fbSend		: FB_SocketSend;(* Send TCP/IP data *)
	fbReceive	: FB_SocketReceive;(* Receive TCP/IP data *)
	nState 		: BYTE;(* Global state *)
	bSndBusy 	: BOOL;(* Tx state *)
	bRcvBusy 	: BOOL;(* Rx state *)
	bDisconnect	: BOOL;(* Disconnect flag, if set the socket will be closed *)

	fbPollTimer	: TON;(* Rx data poll timer *)
	fbResponseTimer	: TON;(* Response timeout timer *)
	fbReconnectTimer : TON;(* Reconnect timer *)

	nS			: UDINT;(* Send frame counter *)
	nR			: UDINT;(* Received frame counter *)
	cbReceived	: UDINT;(* Count of received data bytes *)
	rxBuffer	: ARRAY[0..cTCP_BUFFER_SIZE] OF BYTE;
	cbFrame		: UDINT;(* Rx frame byte size *)
	stTxFrame	: ST_TCPBinaryFrame;(* Tx frame buffer (inclusive header) *)
	stRxFrame	: ST_TCPBinaryFrame;(* Rx frame buffer (inclusive header) *)
	bAbort		: BOOL;(* Flag to abort frame parsing loop *)
	sSend: Tc2_System.T_MaxString;
END_VAR

CASE nState OF
	0:(* Create TCP/IP connection *)
		fbConnect( 	sSrvNetID 		:= sSrvNetID,
					nMode			:= SEL( bLog, 0, CONNECT_MODE_ENABLEDBG ),(* Enable/disable debug output *)
					sRemoteHost 	:= sRemoteHost,
					nRemotePort 	:= nRemotePort,
					tReconnect		:= tReconnect,
					bEnable			:= bEnable,
					eState			=> eState );
		IF NOT fbConnect.bBusy THEN
			IF NOT fbConnect.bError THEN
				IF eState = eSOCKET_CONNECTED THEN(* we are connected *)
					
					fbTx.Clear( sPrefix := CONCAT( sPrefix, 'FB_FrameFifo(sender)::' ), bLog := bLog );(* Clear TX fifo (optional) *)
					fbRx.Clear( sPrefix := CONCAT( sPrefix, 'FB_FrameFifo(receiver)::' ), bLog := bLog );(* Clear RX fifo (optional) *)
					fbLog.Clear( sPrefix := sPrefix, bLog := bLog );(* Clear log fifo (optional) *)
					bSndBusy := FALSE;
					bRcvBusy := FALSE;
					bDisconnect := FALSE;
					cbReceived 	:= 0;(* Reset number of received data bytes *)
					nR 			:= 0;(* Reset receive frame counter *)
					nS 			:= 0;(* Reset send frame counter *)

					fbPollTimer( IN := FALSE, PT := T#0S );
					fbResponseTimer( IN := FALSE, PT := cTCP_RECEIVE_TIMEOUT );
					fbReconnectTimer( IN := FALSE, PT := tReconnect );
				
					fbLog.Message( sMessage := 'Connection established!', hSocket := fbConnect.hSocket );
					nState 	:= 1;
				END_IF
			ELSE(* Connect error => log error *)
				fbLog.Error( sMessage := 'FB_ClientServerConnection()', nErrID := fbConnect.nErrId );
			END_IF
		END_IF


	1:(* Data exchange state *)
		bDisconnect := NOT bEnable OR bDisconnect;(* User/internal disconnect requested? *)
		IF bDisconnect AND NOT bSndBusy AND NOT bRcvBusy THEN
			bDisconnect := FALSE;
			fbLog.Message( sMessage := 'Closing connection!', hSocket := fbConnect.hSocket );
			nState := 2;(* Disconnect *)
		ELSE

			(* --------------------------- Send tx data --------------------------------- *)
			IF NOT bDisconnect AND NOT bSndBusy THEN
				fbTx.RemoveHead();(* Remove oldest user data entry *)
				IF fbTx.bOk THEN(* Success *)
						
					stTxFrame.data := fbTx.stGet;
					
					(* Append/create some protocol header *)
					stTxFrame.head.dwStart 	:= 16#BECF1234;(* Frame start bytes *)
					stTxFrame.head.cbLength := SIZEOF( stTxFrame.data);(* Set length of user data *)
					stTxFrame.head.nS 		:= nS;(* Number of send frames *)
					stTxFrame.head.nR 		:= nR;(* Number of received frames *)
					
					(* Send frame *)
					fbSend( bExecute := FALSE );
// 					sSend := BYTEARR_TO_MAXSTRING(stTxFrame.data);
					
					fbSend(	sSrvNetID 	:= sSrvNetID,
							hSocket		:= fbConnect.hSocket,
							cbLen		:= SIZEOF(TCP_DATA),(* Size of header + size of user data *)
							pSrc		:= ADR(stTxFrame.data),(* Pointer to the frame data *)
							bExecute	:= TRUE );
					bSndBusy := TRUE;
				END_IF
			ELSE(* Wait until send not busy *)
				fbSend( bExecute := FALSE );
				IF NOT fbSend.bBusy THEN
					bSndBusy := FALSE;
					IF NOT fbSend.bError THEN(* No error *)
						nS := nS + 1;(* Increment the number of send frames *)
					ELSE(* Send error => Log error and disconnect *)
						fbLog.Error( sMessage := 'FB_SocketSend()', nErrID := fbSend.nErrId );
						bDisconnect := TRUE;(* Set flag *)
					END_IF
				END_IF
			END_IF
			(* -------------------------------------------------------------------------- *)

// 			(* ------------------ Get/fetch rx data ------------------------------------- *)
// 			IF NOT bDisconnect AND NOT bRcvBusy THEN
// 				fbPollTimer( IN := TRUE );
// 				IF fbPollTimer.Q THEN
// 					IF fbRx.cbFree >= SIZEOF(stRxFrame.data) THEN(* Check free rx fifo space *)
// 						fbPollTimer( IN := FALSE, PT := cTCP_RECEIVE_POLLING_TIME );
// 						fbReceive( bExecute := FALSE );
// 						fbReceive( 	sSrvNetId	:= sSrvNetID,
// 									hSocket		:= fbConnect.hSocket,
// 									cbLen		:= SIZEOF(rxBuffer) - cbReceived,
// 									pDest		:= ADR(rxBuffer) + cbReceived,
// 									bExecute	:= TRUE );
// 						bRcvBusy := TRUE;
// 					END_IF
// 				END_IF
// 				
// 			ELSE(* Wait until receive not busy *)
// 				
// 				fbReceive( bExecute := FALSE );
// 				IF NOT fbReceive.bBusy THEN
// 					bRcvBusy := FALSE;
// 					IF NOT fbReceive.bError THEN
// 						IF fbReceive.nRecBytes > 0 THEN (* Some bytes received *)
// 
// 							fbPollTimer( IN := FALSE, PT := T#0S );(* Bytes received => increase the read (polling) speed *)
// 							fbResponseTimer( IN := FALSE );(* Bytes received => disable timeout check *)
// 							cbReceived := cbReceived + fbReceive.nRecBytes;
// 
// 							(* Parse received bytes *)
// 							REPEAT
// 								bAbort := TRUE;(* Set flag *)
// 								
// 								IF cbReceived >= SIZEOF(stRxFrame.head) THEN (* All header bytes received => check header data *)
// 									
// 									MEMCPY( ADR( stRxFrame.head ), ADR( rxBuffer ), SIZEOF( stRxFrame.head ) );(* Get header data *)
// 								
// 									IF (stRxFrame.head.dwStart = 16#BECF1234) (* Check start bytes *)
// 									AND (stRxFrame.head.nS = nR )(* Check counter (send counter == expected receive counter?) *)
// 									AND (stRxFrame.head.cbLength <= SIZEOF(stRxFrame.data))(* Check frame (user data) length *)
// 									THEN
// 									
// 										cbFrame := SIZEOF(stRxFrame.head) + stRxFrame.head.cbLength;(* Calculate the expected receive frame length *)
// 										IF cbReceived >= cbFrame  THEN (* All frame (user data) bytes received? *)
// 	
// 											MEMCPY( ADR( stRxFrame ), ADR( rxBuffer ), MIN( SIZEOF(stRxFrame), cbFrame ) );
// 											fbRx.AddTail( stPut := stRxFrame.data );(* Add user data to the rx fifo *)
// 											IF fbRx.bOk THEN
// 												nR := nR + 1;(* Increment receive counter *)
// 
// 												MEMMOVE( ADR( rxBuffer ), ADR( rxBuffer ) + cbFrame, cbReceived - cbFrame );(* Shift the remaining rx bytes *)
// 												cbReceived := cbReceived - cbFrame;(* Recalculate the size of the remaining rx bytes *)
// 
// 												IF fbRx.cbFree >= SIZEOF(stRxFrame.data) THEN
// 													bAbort := FALSE;(* reset flag, try to parse next frame *)
// 												END_IF
// 											ELSE (* Fifo overflow => log error and disconnect *)
// 												fbLog.Error( sMessage := 'FB_FrameFifo(receiver)', nErrID := cTCP_ERROR_RECFIFO_OVERFLOW );
// 												bDisconnect := TRUE;(* Set flag *)
// 												RETURN;
// 											END_IF
// 
// (*										ELSE repeat reading *)
// 										END_IF
// 
// 									ELSE(* Receive error => Invalid frame format/data *)
// 										fbLog.Error( sMessage := 'FB_ClientConnection()', nErrID := cTCP_ERROR_INVALID_FRAME_FORMAT );
// 										bDisconnect := TRUE;(* Set flag *)
// 										RETURN;
// 									END_IF
// 
// (*								ELSE repeat reading *)
// 								END_IF (* IF cbReceived >= SIZEOF(stRxFrame.head) THEN *)
// 
// 							UNTIL bAbort
// 							END_REPEAT
// 
// 						ELSE(* No bytes received *)
// 							fbResponseTimer( IN := TRUE );(* No bytes received => enable timeout check *)
// 							IF fbResponseTimer.Q THEN (* Timeout error*)
// 								fbResponseTimer( IN := FALSE );
// 								fbLog.Error( sMessage := 'FB_ClientConnection()', nErrID := cTCP_ERROR_RECEIVE_TIMEOUT );
// 								bDisconnect := TRUE;(* Set flag *)
// 							END_IF							
// 						END_IF(* IF fbReceive.nRecBytes > 0 THEN *)
// 
// 					ELSE(* Receive error => Log error and disconnect *)
// 						fbLog.Error( sMessage := 'FB_SocketReceive()', nErrID := fbReceive.nErrId );
// 						bDisconnect := TRUE;(* set flag *)
// 					END_IF
// 
// 				END_IF(* IF NOT fbReceive.bBusy THEN *)
// 				
// 			END_IF(* IF NOT bDisconnect AND NOT bRcvBusy THEN *)
// 			(* -------------------------------------------------------------------------- *)
			
			
		END_IF(* IF bDisconnect AND NOT bSndBusy AND NOT bRcvBusy THEN *)


	2:(* Disconnect *)
		fbConnect( bEnable:= FALSE, eState=>eState );
		IF eState = eSOCKET_DISCONNECTED THEN
			fbReconnectTimer( IN := TRUE );(* Please wait some seconds and then try to connect again *)
			IF fbReconnectTimer.Q THEN
				fbReconnectTimer( IN := FALSE );
				nState := 0;
			END_IF
		END_IF


END_CASE

END_FUNCTION_BLOCK

// ---- POUs/P_IEC61850_MAIN.TcPOU
PROGRAM P_IEC61850_MAIN
VAR
	fbIEC 	: FB_IEC61850;	
END_VAR

fbIEC();

END_PROGRAM

// ---- POUs/IEC61850Server/FB_IEC61850.TcPOU
FUNCTION_BLOCK FB_IEC61850
VAR
	bInitDone: BOOL := FALSE;	

	i: UDINT;
	j: UDINT;
END_VAR

IF NOT bInitDone THEN
	F_IEC61850ServerInit();

	bInitDone := TRUE;
END_IF

FOR i := 1 TO c_nNumTurbines DO
	fbServer[i].Execute();
	FOR j := 1 TO c_nNumSessions DO
		fbSession[i,j]();
	END_FOR
END_FOR

END_FUNCTION_BLOCK

// ---- POUs/IEC61850Server/F_IEC61850ServerInit.TcPOU
FUNCTION F_IEC61850ServerInit
VAR
	i: UDINT;
	j: UDINT;
END_VAR

FOR i := 1 TO c_nNumTurbines DO
	fbServer[i].ipIED := fbWTURBINE[i];
	
	
	fbServer[i].settings.bEnable := TRUE;
	fbServer[i].settings.sLocalHost := c_aIpAddr;
	fbServer[i].settings.nLocalPort := c_aMMSPortBase + i - 1;
	fbServer[i].settings.sCalled_T_Selector := F_BuildSelector(i);
	fbServer[i].settings.sCalled_S_Selector := F_BuildSelector(i);
	fbServer[i].settings.sCalled_P_Selector := CONCAT('00 00 ', F_UdintToStringPadded(i, 2));
	fbServer[i].settings.sCalled_AP_Title := F_BuildAPTitle(i);
	fbServer[i].settings.nCalled_AP_InvID := i;
	fbServer[i].settings.nCalled_AE_InvID := i;
	fbServer[i].settings.nCalling_AP_InvID := i - 1;
	fbServer[i].settings.nCalling_AE_InvID := i - 1;
	
	FOR j := 1 TO c_nNumSessions DO
		fbSession[i,j].fbConnection.ipServer := fbServer[i];
		fbSession[i,j].fbConnection.settings.bEnable := TRUE;
		fbSession[i,j].nID := i;
	END_FOR
	
	fbWTURBINE[i].WTURBINELD0.WPPD1.ds01.OnInit();
END_FOR

END_FUNCTION

// ---- POUs/IEC61850Server/Util/F_BuildSelector.TcPOU
FUNCTION F_BuildSelector : STRING
VAR_INPUT
    iValue : UDINT;
END_VAR

F_BuildSelector := CONCAT('00 ', F_UdintToStringPadded(iValue, 2));

END_FUNCTION

// ---- POUs/IEC61850Server/Util/F_UdintToStringPadded.TcPOU
FUNCTION F_UdintToStringPadded : STRING
VAR_INPUT
    iValue : UDINT;
    nWidth : DINT;
END_VAR

VAR
    sTemp : STRING(20);
END_VAR

sTemp := UDINT_TO_STRING(iValue);
WHILE LEN(sTemp) < nWidth DO
    sTemp := CONCAT('0', sTemp);
END_WHILE

F_UdintToStringPadded := sTemp;

END_FUNCTION

// ---- POUs/IEC61850Server/Util/F_BuildAPTitle.TcPOU
FUNCTION F_BuildAPTitle : STRING
VAR_INPUT
    iValue : UDINT;
END_VAR

F_BuildAPTitle := CONCAT('1.1.1.999.', UDINT_TO_STRING(iValue));

END_FUNCTION

// ---- POUs/UDP_RX_MAIN.TcPOU
PROGRAM UDP_RX_MAIN
VAR
	fbCloseAll 			: FB_SocketCloseAll;
   	bInitialize			: BOOL := TRUE;
	
	bEnable				: BOOL 			:= TRUE;(* TRUE => Enable/connect, FALSE => Disable/disconnect *)
	bLog				: BOOL			:= TRUE;(* TRUE => Enable log message output, FALSE => Disable *)
	
	fbRx				: FB_UDPRxStateMachine := (sPrefix := 'UDP_RX::');
END_VAR

(* On PLC reset or program download close all opened/created sockets *)
fbCloseAll( sSrvNetId := sSrvNetId, bExecute:= bInitialize );
IF fbCloseAll.bBusy OR fbCloseAll.bError THEN
	RETURN;
END_IF
// IF NOT fbCloseAll.nErrId THEN
//     RETURN; // Not done yet
// END_IF
bInitialize := FALSE;

fbRx(fbRxFifo:=fbRxFIFO, bEnable:=bEnable, bLog:=bLog);

END_PROGRAM

// ---- POUs/UDP/FB_UDPRxStateMachine.TcPOU
FUNCTION_BLOCK FB_UDPRxStateMachine
VAR_IN_OUT
	fbRxFIFO		: FB_UDPFrameFIFO;
END_VAR
VAR_INPUT
	bEnable			: BOOL			:= FALSE;
	tReconnect		: TIME			:= T#5S;
	bLog			: BOOL			:= FALSE;
	sPrefix			: STRING		:= 'UDP_RX::';
END_VAR
VAR_OUTPUT
	bCreated		: BOOL			:= FALSE;
END_VAR
VAR
	fbCreate		: FB_SocketUdpCreate;
	fbClose			: FB_SocketClose;
	hSocket			: T_HSOCKET;
	fbReceiveFrom	: FB_SocketUdpReceiveFrom;
	stReceivedFrom	: ST_UDPFrameEntry;
	fbCreateTimer	: TON := ( PT := T#0S );	
	eState			: E_UDPClientServerState;
END_VAR

CASE eState OF
	(* Idle State *)
	eUDP_STATE_IDLE:
		IF bEnable XOR bCreated THEN
			IF bEnable THEN
				(* Clear rx fifo *)
				fbRxFIFO.Clear( sPrefix := CONCAT( sPrefix, 'FB_FrameFifo(sender)::' ), bLog := bLog );
				
				(* At program start (first time) connect immediately, next time after delay time *)
				fbCreateTimer( IN := TRUE );
				IF fbCreateTimer.Q THEN
					fbCreateTimer( IN := FALSE, PT := tReconnect ); 
					eState := eUDP_STATE_CREATE_START;
				END_IF
			ELSE
				eState := eUDP_STATE_CLOSE_START;
			END_IF
		ELSIF bCreated THEN
			eState := eUDP_STATE_RECEIVE_START;
// 			fbRxFIFO.RemoveHead( stGet => stSendTo );
// 			IF fbRxFIFO.bOk THEN
// 				eState := eUDP_STATE_SEND_START;
// 			END_IF
		ELSE
			fbCreateTimer( IN := FALSE, PT := T#0S );
		END_IF
	
	(* Creation States *)
	eUDP_STATE_CREATE_START:
		fbCreate( bExecute := FALSE  );
		fbCreate( sSrvNetId := sSrvNetId, sLocalHost:= sLocalHost, nLocalPort:= nLocalRxPort, bExecute:= TRUE );
		eState := eUDP_STATE_CREATE_WAIT;

	eUDP_STATE_CREATE_WAIT:
		fbCreate( bExecute := FALSE );
		IF NOT fbCreate.bBusy THEN
			IF NOT fbCreate.bError THEN
				bCreated := TRUE;
				hSocket := fbCreate.hSocket;
// 				fbLog.Message( sMessage := 'Connectionless (UDP) socket created!', hSocket := fbCreate.hSocket );
				eState := eUDP_STATE_IDLE;
			ELSE
// 				fbLog.Error( sMessage := 'FB_SocketUdpCreate()', nErrID := fbCreate.nErrID );
				eState := eUDP_STATE_ERROR;
			END_IF
		END_IF
		
	eUDP_STATE_RECEIVE_START:
		MEMSET( ADR( stReceivedFrom ), 0, SIZEOF( stReceivedFrom ) );
		fbReceiveFrom( bExecute := FALSE );
		fbReceiveFrom( sSrvNetId := sSrvNetId, 
						pDest:= ADR( stReceivedFrom.sMessage ),
						cbLen:= SIZEOF( stReceivedFrom.sMessage ) - 1, (* Without string delimiter *)
						hSocket:= fbCreate.hSocket, bExecute:= TRUE );
		eState := eUDP_STATE_RECEIVE_WAIT;

	eUDP_STATE_RECEIVE_WAIT:
		fbReceiveFrom( bExecute := FALSE );
		IF NOT fbReceiveFrom.bBusy THEN
			IF NOT fbReceiveFrom.bError THEN
				IF fbReceiveFrom.nRecBytes > 0 THEN
					
					stReceivedFrom.stRemoteAddr.sAddr := fbReceiveFrom.sRemoteHost;
					stReceivedFrom.stRemoteAddr.nPort := fbReceiveFrom.nRemotePort;
					
					fbRxFIFO.AddTail( stPut := stReceivedFrom );
	// 				IF NOT fbRxFIFO.bOk THEN(* Check for fifo overflow *)
	// 					fbLog.Error( sMessage :='FB_FrameFifo(receiver)', nErrID := PLCPRJ_ERROR_RECFIFO_OVERFLOW );
	// 				END_IF
				END_IF
				eState := eUDP_STATE_IDLE;
			ELSE
	// 			fbLog.Error( sMessage := 'FB_SocketUdpReceiveFrom()', nErrID := fbReceiveFrom.nErrID );
				IF fbReceiveFrom.nErrID = 16#80072746 THEN(* Connection is reset by remote side *)
					eState := eUDP_STATE_IDLE;
				ELSE
					eState := eUDP_STATE_ERROR;
				END_IF
			END_IF
		END_IF
		
		
	(* Closing States *)
	eUDP_STATE_CLOSE_START:
// 		fbLog.Message( sMessage := 'Closing connectionless (UDP) socket!', hSocket := fbCreate.hSocket );
		fbClose( bExecute := FALSE );
		fbClose( sSrvNetId := sSrvNetId, hSocket := fbCreate.hSocket, bExecute := TRUE );
		eState := eUDP_STATE_CLOSE_WAIT;
		
	eUDP_STATE_CLOSE_WAIT:
		fbClose( bExecute := FALSE );
		IF NOT fbClose.bBusy THEN
			bCreated := FALSE;
			IF NOT fbClose.bError THEN
				eState := eUDP_STATE_IDLE;
			ELSE
// 				fbLog.Error( sMessage := 'FB_SocketClose()', nErrID := fbClose.nErrID );
				eState := eUDP_STATE_ERROR;
			END_IF
		END_IF

	(* Error State *)

	eUDP_STATE_ERROR: (* Error step *)
		IF bCreated THEN
			eState := eUDP_STATE_CLOSE_START;
		ELSE
			eState := eUDP_STATE_IDLE;
		END_IF
		
END_CASE

//FB_Exit must be implemented explicitly. If there is an implementation, then the
//method is called before the controller removes the code of the function block instance
//(implicit call). The return value is not evaluated.
METHOD FB_Exit: BOOL
VAR_INPUT
    bInCopyCode: BOOL;  // TRUE: the exit method is called in order to leave the instance which will be copied afterwards (online change).  
END_VAR
IF bCreated THEN
    fbClose(sSrvNetId := '', hSocket := hSocket, bExecute := TRUE);
END_IF
END_METHOD

END_FUNCTION_BLOCK

// ---- POUs/UDP/Util/FB_UDPFrameFIFO.TcPOU
(* Tx/Rx (string data) fifo control function block *)
FUNCTION_BLOCK FB_UDPFrameFIFO
VAR_INPUT
	bLog		: BOOL := FALSE;(* TRUE => Enable log message output, FALSE => Disable *)
	sPrefix		: STRING := 'Unknown::';(* Log message description string (allows the identification of log message source) *)
	stPut		: ST_UDPFrameEntry;(* Frame entry to add (write) to the buffer *)
END_VAR
VAR_OUTPUT
	bOk			: BOOL;(* TRUE = New entry added or removed succesfully, FALSE = Fifo overflow or fifo empty *)
	stGet		: ST_UDPFrameEntry;(* Frame entry removed (read) from fifo *)
	nCount		: UDINT := 0;(* Number of fifo entries *)
END_VAR
VAR
	fbBuffer 	: FB_MemRingBuffer;(* Basic (lower level) string buffer control function block *)
	buffer		: ARRAY[0..UDP_RX_BUFFER_SIZE] OF BYTE;(* Internal buffer memory *)
	fbCriticalSection:	FB_IecCriticalSection; (* Critical Section required for thread-safety *)
END_VAR

ACTION AddTail:
(* Adds new fifo entry *)
// IF fbCriticalSection.Enter() THEN
	fbBuffer.A_AddTail( pBuffer:= ADR(buffer), cbBuffer:= SIZEOF(buffer),
					pWrite:= ADR( stPut ), cbWrite := SIZEOF( stPut ), 
					bOk=>bOk, nCount=>nCount );
					
// 	fbCriticalSection.Leave();
// END_IF
// IF bOk AND bLog THEN(* Log message *)
// 	ADSLOGSTR( ADSLOG_MSGTYPE_HINT OR ADSLOG_MSGTYPE_LOG, 
// 			CONCAT( CONCAT( sPrefix, SOCKETADDR_TO_STRING(stPut.stRemoteAddr) ), '>>"%s"' ),
// 			stPut.sMessage );
// END_IF
END_ACTION

ACTION Clear:
(* Clears all fifo entries *)
// stGet.sMessage := 0;
// IF fbCriticalSection.Enter() THEN
	MEMSET(ADR(stGet.sMessage), 0, SIZEOF(stGet.sMessage));
	stGet.stRemoteAddr.nPort := 0;
	stGet.stRemoteAddr.sAddr := '';
	fbBuffer.A_Reset( pBuffer := ADR( buffer ), cbBuffer := SIZEOF( buffer ), bOk=>bOk, nCount=>nCount ); 
	
// 	fbCriticalSection.Leave();
// END_IF
END_ACTION

ACTION RemoveHead:
(* Removes oldest fifo entry *)

// IF fbCriticalSection.Enter() THEN
	IF nCount = 0 THEN
		MEMSET(ADR(stGet.sMessage), 0, SIZEOF(stGet.sMessage));
		stGet.stRemoteAddr.nPort := 0;
		stGet.stRemoteAddr.sAddr := '';
		bOk := FALSE;
		RETURN;
	END_IF
	
	fbBuffer.A_RemoveHead( pBuffer:= ADR(buffer), cbBuffer:= SIZEOF(buffer),
							pRead := ADR( stGet ), cbRead := SIZEOF( stGet ),
							bOk=>bOk, nCount=>nCount );
// 	fbCriticalSection.Leave();
// END_IF
END_ACTION

METHOD TEMPRemoveHead : BOOL
VAR_IN_OUT
	stGet	: ST_UDPFrameEntry;
END_VAR
VAR_INPUT
END_VAR
VAR_OUTPUT
	bOk		: BOOL;
END_VAR
IF fbCriticalSection.Enter() THEN
	IF nCount = 0 THEN
		MEMSET(ADR(stGet.sMessage), 0, SIZEOF(stGet.sMessage));
		stGet.stRemoteAddr.nPort := 0;
		stGet.stRemoteAddr.sAddr := '';
		bOk := FALSE;
		RETURN;
	END_IF
	
	fbBuffer.A_RemoveHead( pBuffer:= ADR(buffer), cbBuffer:= SIZEOF(buffer),
							pRead := ADR( stGet ), cbRead := SIZEOF( stGet ),
							bOk=>bOk, nCount=>nCount );
	fbCriticalSection.Leave();
END_IF
END_METHOD

END_FUNCTION_BLOCK

// ---- POUs/UDP_TX_MAIN.TcPOU
PROGRAM UDP_TX_MAIN
VAR
	bSendOnceToRemote	: BOOL;
	bEnable				: BOOL 			:= TRUE;(* TRUE => Enable/connect, FALSE => Disable/disconnect *)
	bLog				: BOOL			:= TRUE;(* TRUE => Enable log message output, FALSE => Disable *)
	
	fbTx				: FB_UDPTxStateMachine := (sPrefix := 'UDP_TX::');
	stSendTo			: ST_UDPFrameEntry;
	
	
	iTemp_1: BYTE := 1;
	iTemp_2: BYTE := 2;
	
	fbCloseAll 			: FB_SocketCloseAll;
	bInitialize: BOOL;
END_VAR

fbCloseAll( sSrvNetId := sSrvNetId, bExecute:= bInitialize );
IF fbCloseAll.bBusy OR fbCloseAll.bError THEN
	RETURN;
END_IF
bInitialize := FALSE;

fbTx(fbTxFifo:=fbTxFIFO, bEnable:=bEnable, bLog:=bLog);

// iTemp_1 := iTemp_1 + 1;
// iTemp_2 := iTemp_2+2;
// 
// IF fbTx.bCreated THEN
// 	IF bSendOnceToRemote THEN
// 		bSendOnceToRemote 			:= FALSE;		(* Clear flag *)
// 		MEMSET(ADR(stSendTo.sMessage), 0, SIZEOF(stSendto.sMessage));
// 		stSendTo.sMessage[1] := INT_TO_BYTE(iTemp_1);
// 		stSendTo.sMessage[2] := INT_TO_BYTE(iTemp_2);		
// 		stSendTo.stRemoteAddr.sAddr := sRemoteHost;	(* Remote host IP address *)
// 		stSendTo.stRemoteAddr.nPort := nRemoteTxPort;	(* Remote host port number *)
// 		fbTxFIFO.AddTail( stPut := stSendTo );	(* Add new entry to the send queue *)
// 	END_IF
// END_IF

END_PROGRAM

// ---- POUs/UDP/FB_UDPTxStateMachine.TcPOU
FUNCTION_BLOCK FB_UDPTxStateMachine
VAR_IN_OUT
	fbTxFIFO		: FB_UDPFrameFIFO;
END_VAR
VAR_INPUT
	bEnable			: BOOL			:= FALSE;			// TRUE => Enable/connect, FALSE => Disable/disconnect
	tReconnect		: TIME			:= T#5S;			// Reconnect delay time
	bLog			: BOOL			:= FALSE;			// TRUE => Enable log message output, FALSE => Disable 
	sPrefix			: STRING 		:= 'PeerToPeerX::'; // Log message description string (allows the identification of log message source)
END_VAR
VAR_OUTPUT
	bCreated		: BOOL;		// Connectionless socket state (TRUE => created, FALSE => closed)
END_VAR
VAR
	fbCreate		: FB_SocketUdpCreate;
	hSocket			: T_HSOCKET;
	fbClose			: FB_SocketClose;
	fbSendTo		: FB_SocketUdpSendTo;
	stSendTo		: ST_UDPFrameEntry;
	fbCreateTimer	: TON := ( PT := T#0S );	
	eState			: E_UDPClientServerState;
END_VAR

CASE eState OF
	(* Idle State *)
	eUDP_STATE_IDLE:
		IF bEnable XOR bCreated THEN
			IF bEnable THEN
				(* Clear send fifo *)
				fbTxFIFO.Clear( sPrefix := CONCAT( sPrefix, 'FB_FrameFifo(sender)::' ), bLog := bLog );
				
				(* At program start (first time) connect immediately, next time after delay time *)
				fbCreateTimer( IN := TRUE );
				IF fbCreateTimer.Q THEN
					fbCreateTimer( IN := FALSE, PT := tReconnect ); 
					eState := eUDP_STATE_CREATE_START;
				END_IF
			ELSE
				eState := eUDP_STATE_CLOSE_START;
			END_IF
		ELSIF bCreated THEN
			fbTxFIFO.RemoveHead( stGet => stSendTo );
			IF fbTxFIFO.bOk THEN
				eState := eUDP_STATE_SEND_START;
			END_IF
		ELSE
			fbCreateTimer( IN := FALSE, PT := T#0S );
		END_IF
	
	(* Creation States *)
	eUDP_STATE_CREATE_START:
		fbCreate( bExecute := FALSE  );
		fbCreate( sSrvNetId := sSrvNetId, sLocalHost:= sLocalHost, nLocalPort:= nLocalTxPort, bExecute:= TRUE );
		eState := eUDP_STATE_CREATE_WAIT;

	eUDP_STATE_CREATE_WAIT:
		fbCreate( bExecute := FALSE );
		IF NOT fbCreate.bBusy THEN
			IF NOT fbCreate.bError THEN
				bCreated := TRUE;
				hSocket := fbCreate.hSocket;
// 				fbLog.Message( sMessage := 'Connectionless (UDP) socket created!', hSocket := fbCreate.hSocket );
				eState := eUDP_STATE_IDLE;
			ELSE
// 				fbLog.Error( sMessage := 'FB_SocketUdpCreate()', nErrID := fbCreate.nErrID );
				eState := eUDP_STATE_ERROR;
			END_IF
		END_IF
	
	(* Sending States *)
	eUDP_STATE_SEND_START:
		fbSendTo( bExecute := FALSE );
		fbSendTo( sSrvNetId := sSrvNetId, sRemoteHost := stSendTo.stRemoteAddr.sAddr,
					nRemotePort := stSendTo.stRemoteAddr.nPort,
					pSrc:= ADR( stSendTo.sMessage ),
					//cbLen:= INT_TO_UDINT(LEN( stSendTo.sMessage )) + 1, (* Include the end delimiter *)
					cbLen := SIZEOF(UDP_DATA),
					hSocket:= fbCreate.hSocket, bExecute:= TRUE );
		eState := eUDP_STATE_SEND_WAIT;

	eUDP_STATE_SEND_WAIT:
		fbSendTo( bExecute := FALSE );
		IF NOT fbSendTo.bBusy THEN
			IF NOT fbSendTo.bError THEN
				eState := eUDP_STATE_IDLE;
			ELSE
// 				fbLog.Error( sMessage := 'FB_SocketUdpSendTo()', nErrID := fbSendTo.nErrID );
				eState := eUDP_STATE_ERROR;
			END_IF
		END_IF
		
	(* Closing States *)
	eUDP_STATE_CLOSE_START:
// 		fbLog.Message( sMessage := 'Closing connectionless (UDP) socket!', hSocket := fbCreate.hSocket );
		fbClose( bExecute := FALSE );
		fbClose( sSrvNetId := sSrvNetId, hSocket := fbCreate.hSocket, bExecute := TRUE );
		eState := eUDP_STATE_CLOSE_WAIT;
		
	eUDP_STATE_CLOSE_WAIT:
		fbClose( bExecute := FALSE );
		IF NOT fbClose.bBusy THEN
			bCreated := FALSE;
			IF NOT fbClose.bError THEN
				eState := eUDP_STATE_IDLE;
			ELSE
// 				fbLog.Error( sMessage := 'FB_SocketClose()', nErrID := fbClose.nErrID );
				eState := eUDP_STATE_ERROR;
			END_IF
		END_IF

	(* Error State *)

	eUDP_STATE_ERROR: (* Error step *)
		IF bCreated THEN
			eState := eUDP_STATE_CLOSE_START;
		ELSE
			eState := eUDP_STATE_IDLE;
		END_IF

END_CASE

//FB_Exit must be implemented explicitly. If there is an implementation, then the
//method is called before the controller removes the code of the function block instance
//(implicit call). The return value is not evaluated.
METHOD FB_Exit: BOOL
VAR_INPUT
    bInCopyCode: BOOL;  // TRUE: the exit method is called in order to leave the instance which will be copied afterwards (online change).  
END_VAR
IF bCreated THEN
    fbClose(sSrvNetId := '', hSocket := hSocket, bExecute := TRUE);
END_IF
END_METHOD

//FB_Init is always available implicitly and it is used primarily for initialization.
//The return value is not evaluated. For a specific influence, you can also declare the
//methods explicitly and provide additional code there with the standard initialization
//code. You can evaluate the return value.
METHOD FB_Init: BOOL
VAR_INPUT
    bInitRetains: BOOL; // TRUE: the retain variables are initialized (reset warm / reset cold)
    bInCopyCode: BOOL;  // TRUE: the instance will be copied to the copy code afterward (online change)   
END_VAR
END_METHOD

END_FUNCTION_BLOCK

// ---- POUs/IEC61850Server/WTURBINE/FB_IED_WTURBINE.TcPOU
{attribute 'no_assign'}
{attribute 'call_after_init'}
FUNCTION_BLOCK FB_IED_WTURBINE EXTENDS FB_AcsiCommonIntelligentElectronicDeviceClass
VAR_INPUT
	WTURBINELD0: FB_LD_WTURBINELD0 := (bLinkResult:=THIS^.AddLogicalDeviceToContainer(ipLogicalDevice:=WTURBINELD0));
END_VAR
VAR
END_VAR

END_FUNCTION_BLOCK

// ---- POUs/IEC61850Server/WTURBINE/LD0/FB_LD_WTURBINELD0.TcPOU
{attribute 'no_assign'}
FUNCTION_BLOCK FB_LD_WTURBINELD0 EXTENDS FB_AcsiCommonLogicalDeviceClass
VAR_INPUT
	LLN0: FB_LN_WTURBINE_LD0_LLN0 := (sClass:='LLN0', bLinkResult:=THIS^.AddLogicalNodeToContainer(ipLogicalNode:=LLN0));
	LPHD1: FB_LN_WTURBINE_LD0_LPHD1 := (sClass:='LPHD', bLinkResult:=THIS^.AddLogicalNodeToContainer(ipLogicalNode:=LPHD1));
	WGEN1: FB_LN_WTURBINE_LD0_WGEN1 := (sClass:='WGEN', bLinkResult:=THIS^.AddLogicalNodeToContainer(ipLogicalNode:=WGEN1));
	WTUR1: FB_LN_WTURBINE_LD0_WTUR1 := (sClass:='WTUR', bLinkResult:=THIS^.AddLogicalNodeToContainer(ipLogicalNode:=WTUR1));
	WROT1: FB_LN_WTURBINE_LD0_WROT1 := (sClass:='WROT', bLinkResult:=THIS^.AddLogicalNodeToContainer(ipLogicalNode:=WROT1));
	WCNV1: FB_LN_WTURBINE_LD0_WCNV1 := (sClass:='WCNV', bLinkResult:=THIS^.AddLogicalNodeToContainer(ipLogicalNode:=WCNV1));
	WMET1: FB_LN_WTURBINE_LD0_WMET1 := (sClass:='WMET', bLinkResult:=THIS^.AddLogicalNodeToContainer(ipLogicalNode:=WMET1));
	WALM1: FB_LN_WTURBINE_LD0_WALM1 := (sClass:='WALM', bLinkResult:=THIS^.AddLogicalNodeToContainer(ipLogicalNode:=WALM1));
	WYAW1: FB_LN_WTURBINE_LD0_WYAW1 := (sClass:='WYAW', bLinkResult:=THIS^.AddLogicalNodeToContainer(ipLogicalNode:=WYAW1));
	WPPD1: FB_LN_WTURBINE_LD0_WPPD1 := (sClass:='WPPD', bLinkResult:=THIS^.AddLogicalNodeToContainer(ipLogicalNode:=WPPD1));
END_VAR
VAR
END_VAR

END_FUNCTION_BLOCK

// ---- POUs/IEC61850Server/WTURBINE/LD0/LLN0/FB_LN_WTURBINE_LD0_LLN0.TcPOU
{attribute 'no_assign'}
FUNCTION_BLOCK FB_LN_WTURBINE_LD0_LLN0 EXTENDS FB_AcsiCommonLogicalNodeClass
VAR_INPUT
	NamPlt: FB_DO_WTURBINE_LD0_LLN0_NamPlt := (sClass:='LPL', bLinkResult:=THIS^.AddDataToContainer(ipData:=NamPlt));
	Beh: FB_DO_WTURBINE_LD0_LLN0_Beh := (sClass:='ENS', bLinkResult:=THIS^.AddDataToContainer(ipData:=Beh));
	Health: FB_DO_WTURBINE_LD0_LLN0_Health := (sClass:='ENS', bLinkResult:=THIS^.AddDataToContainer(ipData:=Health));
	Mod_: FB_DO_WTURBINE_LD0_LLN0_Mod := (sObjectName:='Mod', sClass:='ENC', bLinkResult:=THIS^.AddDataToContainer(ipData:=Mod_));
END_VAR
VAR
END_VAR

END_FUNCTION_BLOCK

// ---- POUs/IEC61850Server/WTURBINE/LD0/LLN0/CDCs/FB_DO_WTURBINE_LD0_LLN0_NamPlt.TcPOU
{attribute 'no_assign'}
FUNCTION_BLOCK FB_DO_WTURBINE_LD0_LLN0_NamPlt EXTENDS FB_AcsiCommonDataClass
VAR_INPUT
	vendor: FB_AcsiDATypeVisString255 := (Fc:=ACSI_FC_DC, bLinkResult:=THIS^.AddDataToContainer(ipData:=vendor));
	swRev: FB_AcsiDATypeVisString255 := (Fc:=ACSI_FC_DC, bLinkResult:=THIS^.AddDataToContainer(ipData:=swRev));
	ldNs: FB_AcsiDATypeVisString255 := (Fc:=ACSI_FC_EX, sValue:='IEC 61850-7-4:2007', bLinkResult:=THIS^.AddDataToContainer(ipData:=ldNs));
END_VAR
VAR
END_VAR

END_FUNCTION_BLOCK

// ---- POUs/IEC61850Server/WTURBINE/LD0/LLN0/CDCs/FB_DO_WTURBINE_LD0_LLN0_Beh.TcPOU
{attribute 'no_assign'}
FUNCTION_BLOCK FB_DO_WTURBINE_LD0_LLN0_Beh EXTENDS FB_AcsiCommonDataClass
VAR_INPUT
	stVal: FB_AcsiDATypeBeh := (Fc:=ACSI_FC_ST, TrgOp:=ACSI_TrgOp_dchg OR ACSI_TrgOp_dupd, bLinkResult:=THIS^.AddDataToContainer(ipData:=stVal));
	q: FB_AcsiDATypeQuality := (Fc:=ACSI_FC_ST, TrgOp:=ACSI_TrgOp_qchg, bLinkResult:=THIS^.AddDataToContainer(ipData:=q));
	t: FB_AcsiDATypeTimeStamp := (Fc:=ACSI_FC_ST, bLinkResult:=THIS^.AddDataToContainer(ipData:=t));
END_VAR
VAR
END_VAR

END_FUNCTION_BLOCK

// ---- POUs/IEC61850Server/WTURBINE/LD0/LLN0/CDCs/FB_DO_WTURBINE_LD0_LLN0_Health.TcPOU
{attribute 'no_assign'}
FUNCTION_BLOCK FB_DO_WTURBINE_LD0_LLN0_Health EXTENDS FB_AcsiCommonDataClass
VAR_INPUT
	stVal: FB_AcsiDATypeHealth := (Fc:=ACSI_FC_ST, TrgOp:=ACSI_TrgOp_dchg OR ACSI_TrgOp_dupd, bLinkResult:=THIS^.AddDataToContainer(ipData:=stVal));
	q: FB_AcsiDATypeQuality := (Fc:=ACSI_FC_ST, TrgOp:=ACSI_TrgOp_qchg, bLinkResult:=THIS^.AddDataToContainer(ipData:=q));
	t: FB_AcsiDATypeTimeStamp := (Fc:=ACSI_FC_ST, bLinkResult:=THIS^.AddDataToContainer(ipData:=t));
END_VAR
VAR
END_VAR

END_FUNCTION_BLOCK

// ---- POUs/IEC61850Server/WTURBINE/LD0/LLN0/CDCs/FB_DO_WTURBINE_LD0_LLN0_Mod.TcPOU
{attribute 'no_assign'}
FUNCTION_BLOCK FB_DO_WTURBINE_LD0_LLN0_Mod EXTENDS FB_AcsiCommonControllableDataClass
VAR_INPUT
	stVal: FB_AcsiDATypeMod := (Fc:=ACSI_FC_ST, TrgOp:=ACSI_TrgOp_dchg, bLinkResult:=THIS^.AddDataToContainer(ipData:=stVal));
	q: FB_AcsiDATypeQuality := (Fc:=ACSI_FC_ST, TrgOp:=ACSI_TrgOp_qchg, bLinkResult:=THIS^.AddDataToContainer(ipData:=q));
	t: FB_AcsiDATypeTimeStamp := (Fc:=ACSI_FC_ST, bLinkResult:=THIS^.AddDataToContainer(ipData:=t));
	ctlModel: FB_AcsiDATypeCtlModels := (Fc:=ACSI_FC_CF, TrgOp:=ACSI_TrgOp_dchg, bLinkResult:=THIS^.AddDataToContainer(ipData:=ctlModel));
	
	fbControl: FB_DirectControl := (ipCtrl:=THIS^.AddServerJob(ipEvent:=fbControl, ipCompletion:=fbControl));
END_VAR
VAR
END_VAR

END_FUNCTION_BLOCK

// ---- POUs/IEC61850Server/FB_DirectControl.TcPOU
FUNCTION_BLOCK FB_DirectControl EXTENDS FB_Control
VAR
	_eControlState: E_DirectControlState; (*State of control state machine*)
END_VAR

METHOD Execute : BOOL
VAR
	bTestOk: BOOL; (*Used to cache the return value of the last '_OperativeTest' or '_DynamicTest' method call*)
	eError: E_AcsiServiceError; (*Used to cache the returned error of the last '_OperativeTest' or '_DynamicTest' method call*)
	tValue: T_UtcTime; (*Used to cache the current system time for 'tOpOk'*)
END_VAR
IF (_ipCtrl <> 0) AND_THEN (_ipCtrl.ipOper <> 0) THEN
	(* Initialize function block in the first cycle *)
	IF NOT bInit THEN
		_Init();
		bInit:=TRUE;
	END_IF

	CASE _eControlState OF
		E_DirectControlState.Ready:
			(* Check if ControlState changed in the last cycle *)
			IF bNewState THEN
				bNewState:=FALSE;
				_Reset();
			END_IF
			(* Check if a valid Oper_req was received *)
			IF bOperReq THEN
				bOperReq:=FALSE;
				(* Go to next ControlState *)
				_eControlState:=E_DirectControlState.PerformTest;
				bNewState:=TRUE;
			END_IF

		E_DirectControlState.PerformTest:
			(* Check if ControlState changed in the last cycle *)
			IF bNewState THEN
				bNewState:=FALSE;
				(* Set 'opRcvd' *)
				IF (_ipCtrl.ipOpRcvd <> 0) THEN
					_ipCtrl.ipOpRcvd.bValue:=TRUE;
				END_IF
			END_IF
			(* Trigger the operative test until it is finished *)
			IF _OperativeTest(bOperativeTestOk=>bTestOk, eError=>eError) THEN
				(* Reset 'opRcvd' *)
				IF (_ipCtrl.ipOpRcvd <> 0) THEN
					_ipCtrl.ipOpRcvd.bValue:=FALSE;
				END_IF
				IF bTestOk THEN
					(* Go to next ControlState *)
					_eControlState:=E_DirectControlState.WaitForExecution;
				ELSE
					fbCompletion.SetCompleted();
					fbCompletion.eServiceError:=eError;
					(* Go back to ControlState 'Ready' *)
					_eControlState:=E_DirectControlState.Ready;
				END_IF
				bNewState:=TRUE;
			END_IF

		E_DirectControlState.WaitForExecution:
			(* Check if ControlState changed in the last cycle *)
			IF bNewState THEN
				bNewState:=FALSE;
			END_IF
			(* Trigger the dynamic test until it is finished *)
			IF _DynamicTest(bDynamicTestOk=>bTestOk, eError=>eError) THEN
				fbCompletion.SetCompleted();
				IF bTestOk THEN
					(* Go to next ControlState *)
					IF (_ipBehVal <> 0) AND_THEN ((_ipBehVal.eValue = E_AcsiBeh.TestBlocked) OR_ELSE (_ipBehVal.eValue = E_AcsiBeh.OnBlocked)) THEN
						_eControlState:=E_DirectControlState.MirrorBlockedCommand;
					ELSE
						_eControlState:=E_DirectControlState.Operate;
					END_IF
				ELSE
					fbCompletion.eServiceError:=eError;
					(* Go back to ControlState 'Ready' *)
					_eControlState:=E_DirectControlState.Ready;
				END_IF
				bNewState:=TRUE;
			END_IF

		E_DirectControlState.Operate:
			(* Check if ControlState changed in the last cycle *)
			IF bNewState THEN
				bNewState:=FALSE;
				(* Set 'opOk' *)
				IF (_ipCtrl.ipOpOk <> 0) THEN
					_ipCtrl.ipOpOk.bValue:=TRUE;
				END_IF
				(* Set 'tOpOk' *)
				IF (_ipCtrl.ipTOpOk <> 0) AND_THEN (_ipCurrentAA <> 0) AND_THEN (_ipCurrentAA.GetSystemTime(tT=>tValue)) THEN
					_ipCtrl.ipTOpOk.tValue:=tValue;
				END_IF
			END_IF
			(* Update value *)
			_SetValue(uCtlVal:=_ipCtrl.ipOper.uCtlVal, ipCtlVal_AV:=_ipCtrl.ipOper.ipCtlVal_AnalogueValue);
			(* Update Timestamp 't' *)
			_UpdateTimestampValue(ipAA:=_ipCurrentAA);

			(* Reset 'opOk' *)
			IF (_ipCtrl.ipOpOk <> 0) THEN
				_ipCtrl.ipOpOk.bValue:=FALSE;
			END_IF
			(* Go back to ControlState 'Ready' *)
			_eControlState:=E_DirectControlState.Ready;
			bNewState:=TRUE;

		E_DirectControlState.MirrorBlockedCommand:
			(* Check if ControlState changed in the last cycle *)
			IF bNewState THEN
				bNewState:=FALSE;
				(* Set 'opOk' *)
				IF (_ipCtrl.ipOpOk <> 0) THEN
					_ipCtrl.ipOpOk.bValue:=TRUE;
				END_IF
				(* Set 'tOpOk' *)
				IF (_ipCtrl.ipTOpOk <> 0) AND_THEN (_ipCurrentAA <> 0) AND_THEN (_ipCurrentAA.GetSystemTime(tT=>tValue)) THEN
					_ipCtrl.ipTOpOk.tValue:=tValue;
				END_IF
			END_IF
			(* Reset 'opOk' *)
			IF (_ipCtrl.ipOpOk <> 0) THEN
				_ipCtrl.ipOpOk.bValue:=FALSE;
			END_IF
			(* Go back to ControlState 'Ready' *)
			_eControlState:=E_DirectControlState.Ready;
			bNewState:=TRUE;
	END_CASE
END_IF

(* Monitor transmission of LastApplError *)
CASE _nLastApplErrorReqState OF
	0:	RETURN;
	1:
		IF (_ipLastApplErrorReq <> 0) THEN
			Execute:=_ipLastApplErrorReq.Execute();
			IF NOT _ipLastApplErrorReq.IsBusy() THEN
				IF _ipLastApplErrorReq.IsCompleted() THEN
					SUPER^.SetCompleted();
				ELSE
					SUPER^.CopyFrom(ipSource:=_ipLastApplErrorReq);
				END_IF
				_nLastApplErrorReqState:=0;
			END_IF
		END_IF
END_CASE
END_METHOD

METHOD OnCompletionWaitEvent : BOOL
VAR_INPUT
	ipDai: I_AcsiDataAccessInfoClass;
	ipData: I_AcsiCommonDataClass;
	eFc: E_AcsiFc;
END_VAR
VAR_OUTPUT
	ipResult: I_AcsiServiceResultClass := fbCompletion;
END_VAR
VAR
	eServiceError: E_AcsiServiceError;
END_VAR
fbCompletion.SetCompleted();
IF (ipDai = 0) OR_ELSE (ipData = 0) THEN
	fbCompletion.eServiceError:=E_AcsiServiceError.AccessViolation;
	RETURN;
END_IF

(* Check if an Operate request is received *)
IF (ipDai.eService = E_AcsiServiceType.SetDataValues) AND_THEN (ipData.sObjectName = 'Oper') THEN
	ScsmAssociation_From_Dai(in:=ipDai, out=>_ipCurrentAA);
	fbCompletion.SetBusy();
	bOperReq:=TRUE;
	OnCompletionWaitEvent:=TRUE;
END_IF
END_METHOD

(*Implementation of user application data update event method.*)
METHOD OnSetVPreEvent : E_AcsiServiceError
VAR_INPUT
	ipDai: I_AcsiDataAccessInfoClass; (*Additional data access info*)
	ipMemory: I_AnyMemoryBuffer; (*Interface pointer to buffer containig new value data*)
	ipData: I_AcsiCommonDataClass; (*Interface pointer to data object*)
	eFc: E_AcsiFc; (*Functional constraint*)
END_VAR
VAR_OUTPUT
	ipLastApplError: I_AcsiDATypeLastApplError; (*IF <> 0 => send LastApplError request*)
END_VAR
VAR
	ipAA: I_ScsmAssociationClass; (*Interface pointer to application association*)
END_VAR
IF (eFc = E_AcsiFc.CO) AND_THEN (_ipCtrl <> 0) AND_THEN (ipDai <> 0) AND_THEN (ipDai.Write) AND_THEN (ipDai.ipAccessData <> 0) AND_THEN ScsmAssociation_From_Dai(in:=ipDai, out=>ipAA) THEN
	IF (_ipCtrl.ipOper <> 0) AND_THEN (_ipCtrl.ipOper.ipOrigin <> 0) AND_THEN (_ipCtrl.ipOper.ipCtlNum <> 0) THEN
		(* Check for invalid write attemps to prevent 'Oper' from being overwritten while a control request is being executed *)
		IF (ipDai.ipAccessData.sObjectName = 'Oper') THEN
			(* Only allow 'Oper' requests in state 'Ready' *)
			IF (_eControlState <> E_DirectControlState.Ready) THEN
				ipLastApplError:=ipAA.SetAdditionalCauseDiag(ipCtrlData:=_ipCtrl.ipOper, eError:=E_AcsiApplError.NoError, stOrigin:=_ipCtrl.ipOper.ipOrigin.stOrigin, nCtlNum:=_ipCtrl.ipOper.ipCtlNum.nValue, eAddCause:=E_AcsiApplAddCause.CommandAlreadyInExecution);
				OnSetVPreEvent:=E_AcsiServiceError.AccessViolation;
			END_IF
		ELSE
			(* Don't allow write access to subdata of 'Oper' *)
			ipLastApplError:=ipAA.SetAdditionalCauseDiag(ipCtrlData:=_ipCtrl.ipOper, eError:=E_AcsiApplError.NoError, stOrigin:=_ipCtrl.ipOper.ipOrigin.stOrigin, nCtlNum:=_ipCtrl.ipOper.ipCtlNum.nValue, eAddCause:=E_AcsiApplAddCause.NotSupported);
			OnSetVPreEvent:=E_AcsiServiceError.AccessViolation;
		END_IF
	END_IF
END_IF
END_METHOD

END_FUNCTION_BLOCK

// ---- POUs/IEC61850Server/FB_Control.TcPOU
FUNCTION_BLOCK FB_Control EXTENDS FB_AsyncServiceResultClass IMPLEMENTS I_AcsiDataAccessEventClass, I_AcsiDataAccessCompletionClass
VAR
	_ipCtrl: I_AcsiCommonControllableDataClass; (* Interface pointer to controllable DO *)
	_eType: E_AcsiCDCType; (* CDC type of the controllable DO *)
	_ipBehVal: I_AcsiDATypeBeh; (* Interface pointer to value of 'Beh' DO of parent LN *)
	_ipStepSize: I_AcsiDATypeAnalogueValue; (* Interface pointer to DO containing stepsize information for BAC *)
	_ipCurrentAA: I_ScsmAssociationClass; (* Interface pointer to association for the current control procedure *)
	_stCurrrentIp: ST_SockAddr; (* IP address of the client for the current control procedure *)
	_ipLastApplErrorReq:  I_AsyncServiceResultClass; (*Interface pointer to LastApplError request service *)
	_nLastApplErrorReqState: BYTE; (* State of LastApplError transmission *)
	_ipCmdTermReq: I_AsyncServiceResultClass; (* Interface pointer to CommandTermination request service *)
	_nCmdTermReqState: BYTE; (* State of CommandTermination transmission *)
	bInit: BOOL; (* Indicates whether this function block has been initialized *)
	bNewState: BOOL; (* Indicates whether the ControlState changed in the last cycle *)
	bOperReq: BOOL; (* Indicates whether a valid Oper_req was received *)
	bSelReq: BOOL; (* Indicates whether a valid Sel_req was received *)
	bSelValReq: BOOL; (* Indicates whether a valid SelVal_req was received *)
	bCancelReq: BOOL; (* Indicates whether a valid Cancel_req was received *)
	fbCompletion: FB_AcsiServiceResultClass; (* Token for CompletionWaitEvent *)
	fbOperCompletion: FB_AcsiServiceResultClass; (* Token for CompletionWaitEvent of Oper_req *)
	fbSelValCompletion: FB_AcsiServiceResultClass; (* Token for CompletionWaitEvent of SelVal_req *)
	fbCancelCompletion: FB_AcsiServiceResultClass; (* Token for CompletionWaitEvent of Cancel_req *)
END_VAR

(* Checks if the value of 'Oper.ctlVal' is valid.
	Return value: TRUE => Value is valid; FALSE => Value is invalid. *)
METHOD PROTECTED _CheckCtlVal : BOOL
VAR_INPUT
	uCtlVal: U_AcsiCtlVal; (* Value of 'ctlVal' DA *)
END_VAR
VAR_OUTPUT
	eError: E_AcsiApplError; (* Error *)
	eAddCause: E_AcsiApplAddCause; (* Application error code *)
END_VAR
VAR
END_VAR
IF (_ipCtrl = 0) OR_ELSE (_eType = E_AcsiCDCType.none) THEN
	RETURN;
END_IF

CASE _eType OF
	E_AcsiCDCType.SPC:
		IF _ipCtrl.ipStVal_BOOLEAN = 0 THEN
			RETURN;
		END_IF
		IF uCtlVal.SPC = _ipCtrl.ipStVal_BOOLEAN.bValue THEN
			eError:= E_AcsiApplError.NoError;
			eAddCause:= E_AcsiApplAddCause.PositionReached;
		ELSE
			_CheckCtlVal:= TRUE;
		END_IF

	E_AcsiCDCType.DPC:
		IF _ipCtrl.ipStVal_Dbpos = 0 THEN
			RETURN;
		END_IF
		IF (SEL(uCtlVal.DPC, E_AcsiDbpos.Off, E_AcsiDbpos.On)) = _ipCtrl.ipStVal_Dbpos.eValue THEN
			eError:= E_AcsiApplError.NoError;
			eAddCause:= E_AcsiApplAddCause.PositionReached;
		ELSE
			_CheckCtlVal:= TRUE;
		END_IF

	E_AcsiCDCType.INC:
		IF _ipCtrl.ipStVal_INT32 = 0 THEN
			RETURN;
		END_IF
		IF uCtlVal.INC = _ipCtrl.ipStVal_INT32.iValue THEN
			eError:= E_AcsiApplError.NoError;
			eAddCause:= E_AcsiApplAddCause.PositionReached;
		ELSE
			_CheckCtlVal:= TRUE;
		END_IF

	E_AcsiCDCType.ENC:
		IF _ipCtrl.ipStVal_ENUMERATED = 0 THEN
			RETURN;
		END_IF
		IF uCtlVal.ENC.iAny = _ipCtrl.ipStVal_ENUMERATED.iAny THEN
			eError:= E_AcsiApplError.NoError;
			eAddCause:= E_AcsiApplAddCause.PositionReached;
		ELSE
			_CheckCtlVal:= TRUE;
		END_IF

	E_AcsiCDCType.BSC:
		IF _ipCtrl.ipValWTr = 0 THEN
			RETURN;
		END_IF
		CASE uCtlVal.BSC OF
			E_AcsiTcmd.Reserved:
				eError:= E_AcsiApplError.NoError;
				eAddCause:= E_AcsiApplAddCause.PositionReached;

			E_AcsiTcmd.Lower:
				IF _ipCtrl.ipValWTr.iPosVal = -64 THEN
					eError:= E_AcsiApplError.NoError;
					eAddCause:= E_AcsiApplAddCause.StepLimit;
				ELSE
					_CheckCtlVal:= TRUE;
				END_IF

			E_AcsiTcmd.Higher:
				IF _ipCtrl.ipValWTr.iPosVal = 63 THEN
					eError:= E_AcsiApplError.NoError;
					eAddCause:= E_AcsiApplAddCause.StepLimit;
				ELSE
					_CheckCtlVal:= TRUE;
				END_IF

			E_AcsiTcmd.Stop:
				_CheckCtlVal:= TRUE;
		END_CASE

	E_AcsiCDCType.ISC:
		IF _ipCtrl.ipValWTr = 0 THEN
			RETURN;
		END_IF
		IF (uCtlVal.ISC < -64) OR_ELSE (uCtlVal.ISC > 63) THEN
			eError:= E_AcsiApplError.NoError;
			eAddCause:= E_AcsiApplAddCause.InconsistentParameters;
		ELSE
			_CheckCtlVal:= TRUE;
		END_IF

	E_AcsiCDCType.APC:
		IF _ipCtrl.ipMxVal = 0 THEN
			RETURN;
		ELSE
			_CheckCtlVal:= TRUE;
		END_IF

	E_AcsiCDCType.BAC:
		IF _ipCtrl.ipMxVal = 0 THEN
			RETURN;
		ELSE
			CASE uCtlVal.BAC OF
				E_AcsiTcmd.Reserved:
					eError:= E_AcsiApplError.NoError;
					eAddCause:= E_AcsiApplAddCause.NotSupported;

				ELSE
					_CheckCtlVal:= TRUE;
			END_CASE
		END_IF
END_CASE
END_METHOD

(* Checks if the values of two 'ctlVal' are equal.
Return value: TRUE => Values are equal; FALSE => Values are unequal. *)
METHOD PROTECTED _CompareCtlVal : BOOL
VAR_INPUT
	uCtlVal1: U_AcsiCtlVal; (* Value of first 'ctlVal' *)
	uCtlVal2: U_AcsiCtlVal; (* Value of second 'ctlVal' *)
END_VAR
VAR
END_VAR
CASE _eType OF
	E_AcsiCDCType.SPC:
		_CompareCtlVal:= uCtlVal1.SPC = uCtlVal2.SPC;

	E_AcsiCDCType.DPC:
		_CompareCtlVal:= uCtlVal1.DPC = uCtlVal2.DPC;

	E_AcsiCDCType.INC:
		_CompareCtlVal:= uCtlVal1.INC = uCtlVal2.INC;

	E_AcsiCDCType.ENC:
		_CompareCtlVal:= uCtlVal1.ENC.iAny = uCtlVal2.ENC.iAny;

	E_AcsiCDCType.BSC:
		_CompareCtlVal:= uCtlVal1.BSC = uCtlVal2.BSC;

	E_AcsiCDCType.ISC:
		_CompareCtlVal:= uCtlVal1.ISC = uCtlVal2.ISC;

	E_AcsiCDCType.APC:
		_CompareCtlVal:= (uCtlVal1.APC.f = uCtlVal2.APC.f) AND_THEN (uCtlVal1.APC.i = uCtlVal2.APC.i);

	E_AcsiCDCType.BAC:
		_CompareCtlVal:= uCtlVal1.BAC = uCtlVal2.BAC;
END_CASE
END_METHOD

(* This method performs the operative test.
Since this test can take multiple PLC cycles, this method is called every cycle, until it returns TRUE. *)
METHOD PROTECTED _DynamicTest : BOOL
VAR_OUTPUT
	bDynamicTestOk: BOOL; (* Indicates whether the dynamic test was successful *)
	eError: E_AcsiServiceError; (* Error code for negative response *)
END_VAR
VAR
END_VAR
bDynamicTestOk:= TRUE;
_DynamicTest:= TRUE;
END_METHOD

(* Initializes the necessary local values. *)
METHOD PROTECTED _Init
VAR
END_VAR
IF _ipCtrl <> 0 THEN
	(* Set '_eType' according to CDC of the controllable data object *)
	IF _ipCtrl.sClass = 'SPC' THEN
		_eType:= E_AcsiCDCType.SPC;
	ELSIF _ipCtrl.sClass = 'DPC' THEN
		_eType:= E_AcsiCDCType.DPC;
	ELSIF _ipCtrl.sClass = 'INC' THEN
		_eType:= E_AcsiCDCType.INC;
	ELSIF _ipCtrl.sClass = 'ENC' THEN
		_eType:= E_AcsiCDCType.ENC;
	ELSIF _ipCtrl.sClass = 'BSC' THEN
		_eType:= E_AcsiCDCType.BSC;
	ELSIF _ipCtrl.sClass = 'ISC' THEN
		_eType:= E_AcsiCDCType.ISC;
	ELSIF _ipCtrl.sClass = 'APC' THEN
		_eType:= E_AcsiCDCType.APC;
	ELSIF _ipCtrl.sClass = 'BAC' THEN
		_eType:= E_AcsiCDCType.BAC;
	END_IF
	(* Get '_ipBehVal' *)
	IF _ipBehVal = 0 THEN
		_ipBehVal:= _ipCtrl.GetBehVal();
	END_IF
END_IF
END_METHOD

(* This method performs the operative test.
Since this test can take multiple PLC cycles, this method is called every cycle, until it returns TRUE. *)
METHOD PROTECTED _OperativeTest : BOOL
VAR_OUTPUT
	bOperativeTestOk: BOOL; (* Indicates whether the operative test was successful *)
	eError: E_AcsiServiceError; (* Error code for negative response *)
END_VAR
VAR
	eApplError: E_AcsiApplError;
	eApplAddCause: E_AcsiApplAddCause;
END_VAR
IF (_ipCtrl <> 0) AND_THEN (_ipCtrl.ipOper <> 0) THEN
	(* Don't allow Oper_req if 'ctlModel' is set to 'status-only' *)
	IF (_ipCtrl.ipCtlModel <> 0) AND_THEN (_ipCtrl.ipCtlModel.eValue = E_AcsiCtlModels.StatusOnly) THEN
		_SendLastApplError(ipAA:=_ipCurrentAA, ipCtrlData:=_ipCtrl.ipOper, eError:=E_AcsiApplError.NoError, ipOrigin:=_ipCtrl.ipOper.ipOrigin, ipCtlNum:=_ipCtrl.ipOper.ipCtlNum, eAddCause:=E_AcsiApplAddCause.Unknown);
		eError:= E_AcsiServiceError.AccessViolation;
		(* Check if Oper_req is valid for current value of 'Beh' *)
	ELSIF (_ipBehVal <> 0) AND_THEN ((_ipBehVal.eValue = E_AcsiBeh.Off) OR_ELSE ((_ipCtrl.ipOper.ipTest <> 0) AND_THEN (_ipCtrl.ipOper.ipTest.bValue <> ((_ipBehVal.eValue = E_AcsiBeh.Test) OR_ELSE (_ipBehVal.eValue = E_AcsiBeh.TestBlocked))))) THEN
		_SendLastApplError(ipAA:=_ipCurrentAA, ipCtrlData:=_ipCtrl.ipOper, eError:=E_AcsiApplError.NoError, ipOrigin:=_ipCtrl.ipOper.ipOrigin, ipCtlNum:=_ipCtrl.ipOper.ipCtlNum, eAddCause:=E_AcsiApplAddCause.BlockedByMode);
		eError:= E_AcsiServiceError.AccessViolation;
		(* Check if 'ctlVal' is valid *)
	ELSIF NOT _CheckCtlVal(uCtlVal:=_ipCtrl.ipOper.uCtlVal, eError=>eApplError, eAddCause=>eApplAddCause) THEN
		_SendLastApplError(ipAA:=_ipCurrentAA, ipCtrlData:=_ipCtrl.ipOper, eError:=eApplError, ipOrigin:=_ipCtrl.ipOper.ipOrigin, ipCtlNum:=_ipCtrl.ipOper.ipCtlNum, eAddCause:=eApplAddCause);
		eError:= E_AcsiServiceError.AccessViolation;
	ELSE (* Oper_req is valid *)
		RemoteAddress_From_ScsmAssociation(in:=_ipCurrentAA, out=>_stCurrrentIp);
		bOperativeTestOk:= TRUE;
	END_IF
END_IF
_OperativeTest:= TRUE;
END_METHOD

(* Resets all local values. *)
METHOD PROTECTED _Reset
VAR
END_VAR
(* Reset local values *)
_ipCurrentAA:= 0;
_stCurrrentIp.sAddr:= '';
_stCurrrentIp.nPort:= 0;
END_METHOD

(* Resets all values of the 'Cancel' DA to their configured initial values. *)
METHOD _ResetCancelValues
VAR
	ipCancel: I_AcsiDATypeCancel; (* Interface pointer to 'Cancel' DA *)
END_VAR
IF (_ipCtrl = 0) OR_ELSE ((ipCancel:=_ipCtrl.ipCancel) = 0) THEN
	RETURN;
END_IF

IF ipCancel.ipCtlVal <> 0 THEN
	ipCancel.uCtlVal:= ipCancel.uCtlVal_Config;
END_IF
IF ipCancel.ipOperTm <> 0 THEN
	ipCancel.ipOperTm.tValue:= ipCancel.ipOperTm.tConfig;
END_IF
IF ipCancel.ipOrigin <> 0 THEN
	ipCancel.ipOrigin.stOrigin:= ipCancel.ipOrigin.stConfig;
END_IF
IF ipCancel.ipCtlNum <> 0 THEN
	ipCancel.ipCtlNum.nValue:= ipCancel.ipCtlNum.nConfig;
END_IF
IF ipCancel.ipT <> 0 THEN
	ipCancel.ipT.tValue:= ipCancel.ipT.tConfig;
END_IF
IF ipCancel.ipTest <> 0 THEN
	ipCancel.ipTest.bValue:= ipCancel.ipTest.bConfig;
END_IF
END_METHOD

(* Resets all values of the 'Oper' DA to their configured initial values. *)
METHOD PROTECTED _ResetOperValues
VAR
	ipOper: I_AcsiDATypeOper; (* Interface pointer to 'Oper' DA *)
END_VAR
IF (_ipCtrl = 0) OR_ELSE ((ipOper:=_ipCtrl.ipOper) = 0) THEN
	RETURN;
END_IF

IF ipOper.ipCtlVal <> 0 THEN
	ipOper.uCtlVal:= ipOper.uCtlVal_Config;
END_IF
IF ipOper.ipOperTm <> 0 THEN
	ipOper.ipOperTm.tValue:= ipOper.ipOperTm.tConfig;
END_IF
IF ipOper.ipOrigin <> 0 THEN
	ipOper.ipOrigin.stOrigin:= ipOper.ipOrigin.stConfig;
END_IF
IF ipOper.ipCtlNum <> 0 THEN
	ipOper.ipCtlNum.nValue:= ipOper.ipCtlNum.nConfig;
END_IF
IF ipOper.ipT <> 0 THEN
	ipOper.ipT.tValue:= ipOper.ipT.tConfig;
END_IF
IF ipOper.ipTest <> 0 THEN
	ipOper.ipTest.bValue:= ipOper.ipTest.bConfig;
END_IF
END_METHOD

(* Resets all values of the 'SBOw' DA to their configured initial values. *)
METHOD PROTECTED _ResetSBOwValues
VAR
	ipSBOw: I_AcsiDATypeSBOw; (* Interface pointer to 'SBOw' DA *)
END_VAR
IF (_ipCtrl = 0) OR_ELSE ((ipSBOw:=_ipCtrl.ipSBOw) = 0) THEN
	RETURN;
END_IF

IF ipSBOw.ipCtlVal <> 0 THEN
	ipSBOw.uCtlVal:= ipSBOw.uCtlVal_Config;
END_IF
IF ipSBOw.ipOperTm <> 0 THEN
	ipSBOw.ipOperTm.tValue:= ipSBOw.ipOperTm.tConfig;
END_IF
IF ipSBOw.ipOrigin <> 0 THEN
	ipSBOw.ipOrigin.stOrigin:= ipSBOw.ipOrigin.stConfig;
END_IF
IF ipSBOw.ipCtlNum <> 0 THEN
	ipSBOw.ipCtlNum.nValue:= ipSBOw.ipCtlNum.nConfig;
END_IF
IF ipSBOw.ipT <> 0 THEN
	ipSBOw.ipT.tValue:= ipSBOw.ipT.tConfig;
END_IF
IF ipSBOw.ipTest <> 0 THEN
	ipSBOw.ipTest.bValue:= ipSBOw.ipTest.bConfig;
END_IF
IF ipSBOw.ipCheck <> 0 THEN
	ipSBOw.ipCheck.eValue:= ipSBOw.ipCheck.eConfig;
END_IF
END_METHOD

(* Sends a negative CommandTermination request. *)
METHOD PROTECTED _SendCommandTerminationReqNeg : BOOL
VAR_INPUT
	ipAA: I_ScsmAssociationClass; (* Interface pointer to application association *)
	ipCtrlData: I_AcsiCommonDataClass; (* Interface pointer to 'Oper', 'Cancel' or 'SBOw' control object, e.g. 'Relay1/XCBR1.CO.Pos.Oper', 'Relay1/CSWI1.CO.Pos.Cancel', 'Relay1/XCBR1.CO.Pos.SBOw' *)
	eError: E_AcsiApplError; (* Error *)
	ipOrigin: I_AcsiDATypeOriginator; (* Interface pointer to 'origin' attribute *)
	ipCtlNum: I_AcsiBATypeINT8U; (* Interface pointer to 'ctlNum' attribute *)
	eAddCause: E_AcsiApplAddCause; (* Application error code *)
END_VAR
VAR
	ipLastApplError: I_AcsiDATypeLastApplError;
END_VAR
IF (ipAA <> 0) AND_THEN (ipCtrlData <> 0) AND_THEN (ipOrigin <> 0) AND_THEN (ipCtlNum <> 0) THEN
	ipLastApplError:= ipAA.SetAdditionalCauseDiag(ipCtrlData:=ipCtrl, eError:=eError, stOrigin:=ipOrigin.stOrigin, nCtlNum:=ipCtlNum.nValue, eAddCause:=eAddCause);
	ipAA.CommandTerminationReq(ipCtrlData:=ipCtrlData, ipLastApplError:=ipLastApplError, ipResult=>_ipCmdTermReq);
	_nCmdTermReqState:= 1;
END_IF
END_METHOD

(* Sends a positive CommandTermination request. *)
METHOD PROTECTED _SendCommandTerminationReqPos : BOOL
VAR_INPUT
	ipAA: I_ScsmAssociationClass; (* Interface pointer to application association *)
	ipCtrlData: I_AcsiCommonDataClass; (* Interface pointer to 'Oper', 'Cancel' or 'SBOw' control object, e.g. 'Relay1/XCBR1.CO.Pos.Oper', 'Relay1/CSWI1.CO.Pos.Cancel', 'Relay1/XCBR1.CO.Pos.SBOw' *)
END_VAR
VAR
END_VAR
IF (ipAA <> 0) AND_THEN (ipCtrlData <> 0) THEN
	_SendCommandTerminationReqPos:= ipAA.CommandTerminationReq(ipCtrlData:=ipCtrlData, ipLastApplError:=0, ipResult=>_ipCmdTermReq);
	_nCmdTermReqState:= 1;
END_IF
END_METHOD

(* Sends a LastApplError request. *)
METHOD PROTECTED _SendLastApplError : BOOL
VAR_INPUT
	ipAA: I_ScsmAssociationClass; (* Interface pointer to application association *)
	ipCtrlData: I_AcsiCommonDataClass; (* Interface pointer to 'Oper', 'Cancel' or 'SBOw' control object *)
	eError: E_AcsiApplError; (* Error *)
	ipOrigin: I_AcsiDATypeOriginator; (* Interface pointer to 'origin' attribute *)
	ipCtlNum: I_AcsiBATypeINT8U; (* Interface pointer to 'ctlNum' attribute *)
	eAddCause: E_AcsiApplAddCause; (* Application error code *)
END_VAR
VAR
	ipLastApplError: I_AcsiDATypeLastApplError; (* Interface pointer to AdditionalCauseDiag object *)
END_VAR
(* Get values from 'Oper' and send LastApplError *)
IF (ipAA <> 0) AND_THEN (ipOrigin <> 0) AND_THEN (ipCtlNum <> 0) THEN
	ipLastApplError:= ipAA.SetAdditionalCauseDiag(ipCtrlData:=ipCtrlData, eError:=eError, stOrigin:=ipOrigin.stOrigin, nCtlNum:=ipCtlNum.nValue, eAddCause:=eAddCause);

	_SendLastApplError:= ipAA.LastApplErrorReq(ipLastApplError:=ipLastApplError, ipResult=>_ipLastApplErrorReq);
	SUPER^.SetBusy();
	_nLastApplErrorReqState:= 1;
END_IF
END_METHOD

(* Sets the value of 'mxVal' to the value of 'ctlVal'.
Return value: TRUE => Success; FALSE => Failure. *)
METHOD PROTECTED _SetApcValue : BOOL
VAR_INPUT
	ipMxVal: I_AcsiDATypeAnalogueValue; (* Interface pointer to DA that will be written *)
	uCtlVal: U_AcsiCtlVal; (* Value of 'ctlVal' DA *)
	ipCtlVal_AV: I_AcsiDATypeAnalogueValue; (* Interface pointer to 'ctlVal' of type AnalogueValue *)
END_VAR
VAR
END_VAR
IF ((ipMxVal = 0) OR_ELSE ((ipMxVal.ipF = 0) AND_THEN (ipMxVal.ipI = 0))) OR_ELSE ((ipCtlVal_AV = 0) OR_ELSE ((ipCtlVal_AV.ipF = 0) AND_THEN (ipCtlVal_AV.ipI = 0))) THEN
	RETURN;
END_IF

IF ipMxVal.ipF <> 0 THEN
	IF ipCtlVal_AV.ipF <> 0 THEN
		ipMxVal.fValue:= uCtlVal.APC.f;
	ELSE
		(* 'ctlVal.i' is present, but not 'ctlVal.f' -> convert and use value of 'ctlVal.i' *)
		ipMxVal.fValue:= DINT_TO_REAL(uCtlVal.APC.i);
	END_IF
END_IF
IF ipMxVal.ipI <> 0 THEN
	IF ipCtlVal_AV.ipI <> 0 THEN
		ipMxVal.iValue:= uCtlVal.APC.i;
	ELSE
		(* 'ctlVal.if' is present, but not 'ctlVal.i' -> convert and use value of 'ctlVal.f' *)
		ipMxVal.iValue:= REAL_TO_DINT(uCtlVal.APC.f);
	END_IF
END_IF
END_METHOD

(* Increments or decrements the value of 'mxVal' according to the value of 'ctlVal' and 'stepSize'.
If 'stepSize' is not specified, the value 1 is used.
Return value: TRUE => Success; FALSE => Failure. *)
METHOD PROTECTED _SetBacValue : BOOL
VAR_INPUT
	ipMxVal: I_AcsiDATypeAnalogueValue; (* Interface pointer to DA that will be written *)
	uCtlVal: U_AcsiCtlVal; (* Value of 'ctlVal' DA *)
	ipStepSize: I_AcsiDATypeAnalogueValue; (* Interface pointer to 'stepSize' DA (Optional) *)
END_VAR
VAR
	fStepSize: REAL := 1; (* stepSize for 'f' *)
	iStepSize: DINT := 1; (* stepSize for 'i' *)
END_VAR
IF (ipMxVal = 0) OR_ELSE ((ipMxVal.ipF = 0) AND_THEN (ipMxVal.ipI = 0)) THEN
	RETURN;
END_IF

IF (ipStepSize <> 0) AND_THEN (((ipStepSize.ipF <> 0) AND_THEN (ipStepSize.fValue <> 0.0)) OR_ELSE ((ipStepSize.ipI <> 0) AND_THEN (ipStepSize.iValue <> 0))) THEN
	IF ipStepSize.ipF <> 0 THEN
		fStepSize:= ipStepSize.fValue;
	ELSE
		(* 'stepSize.i' is present, but not 'stepSize.f' -> convert and use value of 'stepSize.i' *)
		fStepSize:= DINT_TO_REAL(ipStepSize.iValue);
	END_IF
	IF ipStepSize.ipI <> 0 THEN
		iStepSize:= ipStepSize.iValue;
	ELSE
		(* 'stepSize.f' is present, but not 'stepSize.i' -> convert and use value of 'stepSize.f' *)
		iStepSize:= REAL_TO_DINT(ipStepSize.fValue);
	END_IF
END_IF

CASE uCtlVal.BAC OF
	E_AcsiTcmd.Stop:
		_SetBacValue:= TRUE;

	E_AcsiTcmd.Lower:
		IF ipMxVal.ipF <> 0 THEN
			ipMxVal.fValue:= ipMxVal.fValue - fStepSize;
		END_IF
		IF ipMxVal.ipI <> 0 THEN
			ipMxVal.iValue:= ipMxVal.iValue - iStepSize;
		END_IF
		_SetBacValue:= TRUE;

	E_AcsiTcmd.Higher:
		IF ipMxVal.ipF <> 0 THEN
			ipMxVal.fValue:= ipMxVal.fValue + fStepSize;
		END_IF
		IF ipMxVal.ipI <> 0 THEN
			ipMxVal.iValue:= ipMxVal.iValue + iStepSize;
		END_IF
		_SetBacValue:= TRUE;
END_CASE
END_METHOD

(* Increments or decrements the value of 'valWTr' according to the value of 'ctlVal'.
Return value: TRUE => Success; FALSE => Failure. *)
METHOD PROTECTED _SetBscValue : BOOL
VAR_INPUT
	ipValWTr: I_AcsiDATypeValWithTrans; (* Interface pointer to DA that will be written *)
	uCtlVal: U_AcsiCtlVal; (* Value of 'ctlVal' DA *)
END_VAR
VAR
END_VAR
IF ipValWTr = 0 THEN
	RETURN;
END_IF

CASE uCtlVal.BSC OF
	E_AcsiTcmd.Stop:
		_SetBscValue:= TRUE;

	E_AcsiTcmd.Lower:
		ipValWTr.iPosVal:= ipValWTr.iPosVal - 1;
		_SetBscValue:= TRUE;

	E_AcsiTcmd.Higher:
		ipValWTr.iPosVal:= ipValWTr.iPosVal + 1;
		_SetBscValue:= TRUE;
END_CASE
END_METHOD

(* Sets the value of 'stVal' according to the value of 'ctlVal'.
Return value: TRUE => Success; FALSE => Failure. *)
METHOD PROTECTED _SetDpcValue : BOOL
VAR_INPUT
	ipStVal: I_AcsiDATypeDbpos; (* Interface pointer to DA that will be written *)
	uCtlVal: U_AcsiCtlVal; (* Value of 'ctlVal' DA *)
END_VAR
VAR
END_VAR
IF ipStVal = 0 THEN
	RETURN;
END_IF

ipStVal.eValue:= SEL(uCtlVal.DPC, E_AcsiDbpos.Off, E_AcsiDbpos.On);
_SetDpcValue:= TRUE;
END_METHOD

(* Sets the value of 'stVal' according to the value of 'ctlVal'.
Return value: TRUE => Success; FALSE => Failure. *)
METHOD PROTECTED _SetEncValue : BOOL
VAR_INPUT
	ipStVal: I_AcsiBATypeENUMERATED; (* Interface pointer to DA that will be written *)
	uCtlVal: U_AcsiCtlVal; (* Value of 'ctlVal' DA *)
END_VAR
VAR
END_VAR
IF ipStVal = 0 THEN
	RETURN;
END_IF

ipStVal.iAny:= uCtlVal.ENC.iAny;
_SetEncValue:= TRUE;
END_METHOD

(* Sets the value of 'stVal' to the value of 'ctlVal'.
Return value: TRUE => Success; FALSE => Failure. *)
METHOD PROTECTED _SetIncValue : BOOL
VAR_INPUT
	ipStVal: I_AcsiBATypeINT32; (* Interface pointer to DA that will be written *)
	uCtlVal: U_AcsiCtlVal; (* Value of 'ctlVal' DA *)
END_VAR
VAR
END_VAR
IF ipStVal = 0 THEN
	RETURN;
END_IF

ipStVal.iValue:= uCtlVal.INC;
_SetIncValue:= TRUE;
END_METHOD

(* Sets the value of 'valWTr' to the value of 'ctlVal'.
Return value: TRUE => Success; FALSE => Failure. *)
METHOD PROTECTED _SetIscValue : BOOL
VAR_INPUT
	ipValWTr: I_AcsiDATypeValWithTrans; (* Interface pointer to DA that will be written *)
	uCtlVal: U_AcsiCtlVal; (* Value of 'ctlVal' DA *)
END_VAR
VAR
END_VAR
IF ipValWTr = 0 THEN
	RETURN;
END_IF

ipValWTr.iPosVal:= uCtlVal.ISC;
_SetIscValue:= TRUE;
END_METHOD

(* Sets the value of 'stVal' to the value of 'ctlVal'.
Return value: TRUE => Success; FALSE => Failure. *)
METHOD PROTECTED _SetSpcValue : BOOL
VAR_INPUT
	ipStVal: I_AcsiBATypeBOOLEAN; (* Interface pointer to DA that will be written *)
	uCtlVal: U_AcsiCtlVal; (* Value of 'ctlVal' DA *)
END_VAR
VAR
END_VAR
IF ipStVal = 0 THEN
	RETURN;
END_IF

ipStVal.bValue:= uCtlVal.SPC;
_SetSpcValue:= TRUE;
END_METHOD

(* Sets the value of the respective DA according to the value of 'Oper.ctlVal'.
Return value: TRUE => Success, FALSE => Failure. *)
METHOD PROTECTED _SetValue : BOOL
VAR_INPUT
	uCtlVal: U_AcsiCtlVal; (* Value of 'ctlVal' DA *)
	ipCtlVal_AV: I_AcsiDATypeAnalogueValue; (* Interface pointer to 'ctlVal' of type AnalogueValue *)
END_VAR
VAR
END_VAR
IF _ipCtrl = 0 THEN
	RETURN;
END_IF

CASE _eType OF
	E_AcsiCDCType.SPC:
		_SetValue:= _SetSpcValue(ipStVal:=_ipCtrl.ipStVal_BOOLEAN, uCtlVal:=uCtlVal);

	E_AcsiCDCType.DPC:
		_SetValue:= _SetDpcValue(ipStVal:=_ipCtrl.ipStVal_Dbpos, uCtlVal:=uCtlVal);

	E_AcsiCDCType.INC:
		_SetValue:= _SetIncValue(ipStVal:=_ipCtrl.ipStVal_INT32, uCtlVal:=uCtlVal);

	E_AcsiCDCType.ENC:
		_SetValue:= _SetEncValue(ipStVal:=_ipCtrl.ipStVal_ENUMERATED, uCtlVal:=uCtlVal);

	E_AcsiCDCType.BSC:
		_SetValue:= _SetBscValue(ipValWTr:=_ipCtrl.ipValWTr, uCtlVal:=uCtlVal);

	E_AcsiCDCType.ISC:
		_SetValue:= _SetIscValue(ipValWTr:=_ipCtrl.ipValWTr, uCtlVal:=uCtlVal);

	E_AcsiCDCType.APC:
		_SetValue:= _SetApcValue(ipMxVal:=_ipCtrl.ipMxVal, uCtlVal:=uCtlVal, ipCtlVal_AV:=ipCtlVal_AV);

	E_AcsiCDCType.BAC:
		_SetValue:= _SetBacValue(ipMxVal:=_ipCtrl.ipMxVal, uCtlVal:=uCtlVal, ipStepSize:=_ipStepSize);

END_CASE
END_METHOD

(* This method performs the test of the SelectWithValue operation.
Since this test can take multiple PLC cycles, this method is called every cycle, until it returns TRUE. *)
METHOD PROTECTED _Test : BOOL
VAR_OUTPUT
	bTestOk: BOOL; (* Indicates whether the test was successful *)
	eError: E_AcsiServiceError; (* Error code for negative response *)
END_VAR
VAR
	eApplError: E_AcsiApplError; (* Error *)
	eApplAddCause: E_AcsiApplAddCause; (* Application error code *)
END_VAR
IF (_ipCtrl <> 0) AND_THEN (_ipCtrl.ipSBOw <> 0) THEN
	(* Don't allow control if 'ctlModel' is set to 'status-only' *)
	IF (_ipCtrl.ipCtlModel <> 0) AND_THEN (_ipCtrl.ipCtlModel.eValue = E_AcsiCtlModels.StatusOnly) THEN
		_SendLastApplError(ipAA:=_ipCurrentAA, ipCtrlData:=_ipCtrl.ipSBOw, eError:=E_AcsiApplError.NoError, ipOrigin:=_ipCtrl.ipSBOw.ipOrigin, ipCtlNum:=_ipCtrl.ipSBOw.ipCtlNum, eAddCause:=E_AcsiApplAddCause.Unknown);
		eError:= E_AcsiServiceError.AccessViolation;
		(* Check if 'ctlVal' is valid *)
	ELSIF NOT _CheckCtlVal(uCtlVal:=_ipCtrl.ipSBOw.uCtlVal, eError=>eApplError, eAddCause=>eApplAddCause) THEN
		_SendLastApplError(ipAA:=_ipCurrentAA, ipCtrlData:=_ipCtrl.ipSBOw, eError:=eApplError, ipOrigin:=_ipCtrl.ipSBOw.ipOrigin, ipCtlNum:=_ipCtrl.ipSBOw.ipCtlNum, eAddCause:=eApplAddCause);
		eError:= E_AcsiServiceError.AccessViolation;
		(* SelVal_req is valid *)
	ELSE
		RemoteAddress_From_ScsmAssociation(in:=_ipCurrentAA, out=>_stCurrrentIp);
		bTestOk:= TRUE;
	END_IF
END_IF
_Test:= TRUE;
END_METHOD

(* Sets the value of 't' to the current time.
Return value: TRUE => Success; FALSE => Failure. *)
METHOD PROTECTED _UpdateTimestampValue : BOOL
VAR_INPUT
	ipAA: I_ScsmAssociationClass; (* Interface pointer to application association *)
END_VAR
VAR
	tValue: T_UtcTime; (* Current time *)
END_VAR
IF (ipAA <> 0) AND_THEN (_ipCtrl <> 0) AND_THEN (_ipCtrl.ipT <> 0) THEN
	_UpdateTimestampValue:= ipAA.GetSystemTime(tT=>tValue);
	_ipCtrl.ipT.tValue:= tValue;
END_IF
END_METHOD

PROPERTY eType : E_AcsiCDCType
GET
eType:= _eType;
END_GET
SET
_eType:= eType;
END_SET
END_PROPERTY

PROPERTY ipBehVal : I_AcsiDATypeBeh
GET
ipBehVal:= _ipBehVal;
END_GET
SET
_ipBehVal:= ipBehVal;
END_SET
END_PROPERTY

PROPERTY ipCtrl : I_AcsiCommonControllableDataClass
GET
ipCtrl:= _ipCtrl;
END_GET
SET
_ipCtrl:= ipCtrl;
END_SET
END_PROPERTY

PROPERTY ipStepSize : I_AcsiDATypeAnalogueValue
GET
ipStepSize:= _ipStepSize;
END_GET
SET
_ipStepSize:= ipStepSize;
END_SET
END_PROPERTY

METHOD OnAbort : BOOL
VAR_INPUT
	ipReason: I_ServiceErrorClass;
END_VAR
VAR_OUTPUT
	ipResult: I_AsyncServiceResultClass := THIS^;
END_VAR
VAR
END_VAR
(* Forward Abort to LastApplError request service *)
IF (_ipLastApplErrorReq <> 0) AND_THEN (_ipLastApplErrorReq.IsBusy()) THEN
	_ipLastApplErrorReq.OnAbort(ipReason:=ipReason);
END_IF
(* Forward Abort to CommandTermination request service *)
IF (_ipCmdTermReq <> 0) AND_THEN (_ipCmdTermReq.IsBusy()) THEN
	_ipCmdTermReq.OnAbort(ipReason:=ipReason);
END_IF

SUPER^.SetCompleted();
fbCompletion.SetCompleted();
END_METHOD

METHOD OnCompletionWaitEvent : BOOL
VAR_INPUT
	ipDai: I_AcsiDataAccessInfoClass;
	ipData: I_AcsiCommonDataClass;
	eFc: E_AcsiFc;
END_VAR
VAR_OUTPUT
	ipResult: I_AcsiServiceResultClass := fbCompletion;
END_VAR
VAR
END_VAR
END_METHOD

(* Implementation of user application data update event method. *)
METHOD OnGetVEvent
VAR_INPUT
	ipDai: I_AcsiDataAccessInfoClass; (* Additional data access info *)
	ipData: I_AcsiCommonDataClass; (* Interface pointer to data object *)
	eFc: E_AcsiFc; (* Functional constraint *)
END_VAR
VAR
END_VAR
END_METHOD

(* Implementation of user application data update event method. *)
METHOD OnGetVPreEvent : E_AcsiServiceError
VAR_INPUT
	ipDai: I_AcsiDataAccessInfoClass; (* Additional data access info *)
	ipData: I_AcsiCommonDataClass; (* Interface pointer to data object *)
	eFc: E_AcsiFc; (* Functional constraint *)
END_VAR
VAR
END_VAR
END_METHOD

(* Implementation of user application data update event method. *)
METHOD OnSetVEvent
VAR_INPUT
	ipDai: I_AcsiDataAccessInfoClass; (* Additional data access info *)
	ipData: I_AcsiCommonDataClass; (* Interface pointer to data object *)
	eFc: E_AcsiFc; (* Functional constraint *)
END_VAR
VAR
END_VAR
END_METHOD

(* Implementation of user application data update event method. *)
METHOD OnSetVPreEvent : E_AcsiServiceError
VAR_INPUT
	ipDai: I_AcsiDataAccessInfoClass; (* Additional data access info *)
	ipMemory: I_AnyMemoryBuffer; (* Interface pointer to buffer containig new value data *)
	ipData: I_AcsiCommonDataClass; (* Interface pointer to data object *)
	eFc: E_AcsiFc; (* Functional constraint *)
END_VAR
VAR_OUTPUT
	ipLastApplError: I_AcsiDATypeLastApplError; (* IF <> 0 => send LastApplError request *)
END_VAR
VAR
END_VAR
END_METHOD

END_FUNCTION_BLOCK

// ---- POUs/IEC61850Server/WTURBINE/LD0/LPHD1/FB_LN_WTURBINE_LD0_LPHD1.TcPOU
{attribute 'no_assign'}
FUNCTION_BLOCK FB_LN_WTURBINE_LD0_LPHD1 EXTENDS FB_AcsiCommonLogicalNodeClass
VAR_INPUT
	PhyNam: FB_DO_WTURBINE_LD0_LPHD1_PhyNam := (sClass:='WDPL', bLinkResult:=THIS^.AddDataToContainer(ipData:=PhyNam));
	PhyHealth: FB_DO_WTURBINE_LD0_LPHD1_PhyHealth := (sClass:='ENS', bLinkResult:=THIS^.AddDataToContainer(ipData:=PhyHealth));
	Proxy: FB_DO_WTURBINE_LD0_LPHD1_Proxy := (sClass:='SPS', bLinkResult:=THIS^.AddDataToContainer(ipData:=Proxy));
END_VAR
VAR
END_VAR

END_FUNCTION_BLOCK

// ---- POUs/IEC61850Server/WTURBINE/LD0/LPHD1/CDCs/FB_DO_WTURBINE_LD0_LPHD1_PhyNam.TcPOU
{attribute 'no_assign'}
FUNCTION_BLOCK FB_DO_WTURBINE_LD0_LPHD1_PhyNam EXTENDS FB_AcsiCommonDataClass
VAR_INPUT
	vendor: FB_AcsiDATypeVisString255 := (Fc:=ACSI_FC_DC, bLinkResult:=THIS^.AddDataToContainer(ipData:=vendor));
END_VAR
VAR
END_VAR

END_FUNCTION_BLOCK

// ---- POUs/IEC61850Server/WTURBINE/LD0/LPHD1/CDCs/FB_DO_WTURBINE_LD0_LPHD1_PhyHealth.TcPOU
{attribute 'no_assign'}
FUNCTION_BLOCK FB_DO_WTURBINE_LD0_LPHD1_PhyHealth EXTENDS FB_AcsiCommonDataClass
VAR_INPUT
	stVal: FB_AcsiDATypePhyHealth := (Fc:=ACSI_FC_ST, TrgOp:=ACSI_TrgOp_dchg OR ACSI_TrgOp_dupd, bLinkResult:=THIS^.AddDataToContainer(ipData:=stVal));
	q: FB_AcsiDATypeQuality := (Fc:=ACSI_FC_ST, TrgOp:=ACSI_TrgOp_qchg, bLinkResult:=THIS^.AddDataToContainer(ipData:=q));
	t: FB_AcsiDATypeTimeStamp := (Fc:=ACSI_FC_ST, bLinkResult:=THIS^.AddDataToContainer(ipData:=t));
END_VAR
VAR
END_VAR

END_FUNCTION_BLOCK

// ---- POUs/IEC61850Server/WTURBINE/LD0/LPHD1/CDCs/FB_DO_WTURBINE_LD0_LPHD1_Proxy.TcPOU
{attribute 'no_assign'}
FUNCTION_BLOCK FB_DO_WTURBINE_LD0_LPHD1_Proxy EXTENDS FB_AcsiCommonDataClass
VAR_INPUT
	stVal: FB_AcsiBATypeBOOLEAN := (Fc:=ACSI_FC_ST, TrgOp:=ACSI_TrgOp_dchg, bLinkResult:=THIS^.AddDataToContainer(ipData:=stVal));
	q: FB_AcsiDATypeQuality := (Fc:=ACSI_FC_ST, TrgOp:=ACSI_TrgOp_qchg, bLinkResult:=THIS^.AddDataToContainer(ipData:=q));
	t: FB_AcsiDATypeTimeStamp := (Fc:=ACSI_FC_ST, bLinkResult:=THIS^.AddDataToContainer(ipData:=t));
END_VAR
VAR
END_VAR

END_FUNCTION_BLOCK

// ---- POUs/IEC61850Server/WTURBINE/LD0/WGEN1/FB_LN_WTURBINE_LD0_WGEN1.TcPOU
{attribute 'no_assign'}
FUNCTION_BLOCK FB_LN_WTURBINE_LD0_WGEN1 EXTENDS FB_AcsiCommonLogicalNodeClass
VAR_INPUT
	Beh: FB_DO_WTURBINE_LD0_WGEN1_Beh := (sClass:='ENS', bLinkResult:=THIS^.AddDataToContainer(ipData:=Beh));
	RotSpd: FB_DO_WTURBINE_LD0_WGEN1_RotSpd := (sClass:='MV', bLinkResult:=THIS^.AddDataToContainer(ipData:=RotSpd));
END_VAR
VAR
END_VAR

END_FUNCTION_BLOCK

// ---- POUs/IEC61850Server/WTURBINE/LD0/WGEN1/CDCs/FB_DO_WTURBINE_LD0_WGEN1_Beh.TcPOU
{attribute 'no_assign'}
FUNCTION_BLOCK FB_DO_WTURBINE_LD0_WGEN1_Beh EXTENDS FB_AcsiCommonDataClass
VAR_INPUT
	stVal: FB_AcsiDATypeBeh := (Fc:=ACSI_FC_ST, TrgOp:=ACSI_TrgOp_dchg OR ACSI_TrgOp_dupd, bLinkResult:=THIS^.AddDataToContainer(ipData:=stVal));
	q: FB_AcsiDATypeQuality := (Fc:=ACSI_FC_ST, TrgOp:=ACSI_TrgOp_qchg, bLinkResult:=THIS^.AddDataToContainer(ipData:=q));
	t: FB_AcsiDATypeTimeStamp := (Fc:=ACSI_FC_ST, bLinkResult:=THIS^.AddDataToContainer(ipData:=t));
END_VAR
VAR
END_VAR

END_FUNCTION_BLOCK

// ---- POUs/IEC61850Server/WTURBINE/LD0/WGEN1/CDCs/FB_DO_WTURBINE_LD0_WGEN1_RotSpd.TcPOU
{attribute 'no_assign'}
FUNCTION_BLOCK FB_DO_WTURBINE_LD0_WGEN1_RotSpd EXTENDS FB_AcsiCommonDataClass
VAR_INPUT
	mag: FB_AcsiDATypeAnalogueValue := (Fc:=ACSI_FC_MX, TrgOp:=ACSI_TrgOp_dchg OR ACSI_TrgOp_dupd, i:=(bPresence:=FALSE), bLinkResult:=THIS^.AddDataToContainer(ipData:=mag));
	q: FB_AcsiDATypeQuality := (Fc:=ACSI_FC_MX, TrgOp:=ACSI_TrgOp_qchg, bLinkResult:=THIS^.AddDataToContainer(ipData:=q));
	t: FB_AcsiDATypeTimeStamp := (Fc:=ACSI_FC_MX, bLinkResult:=THIS^.AddDataToContainer(ipData:=t));
END_VAR
VAR
END_VAR

END_FUNCTION_BLOCK

// ---- POUs/IEC61850Server/WTURBINE/LD0/WTUR1/FB_LN_WTURBINE_LD0_WTUR1.TcPOU
{attribute 'no_assign'}
FUNCTION_BLOCK FB_LN_WTURBINE_LD0_WTUR1 EXTENDS FB_AcsiCommonLogicalNodeClass
VAR_INPUT
	Beh: FB_DO_WTURBINE_LD0_WTUR1_Beh := (sClass:='ENS', bLinkResult:=THIS^.AddDataToContainer(ipData:=Beh));
	TotWh: FB_DO_WTURBINE_LD0_WTUR1_TotWh := (sClass:='CTE', bLinkResult:=THIS^.AddDataToContainer(ipData:=TotWh));
	TurSt: FB_DO_WTURBINE_LD0_WTUR1_TurSt := (sClass:='STV', bLinkResult:=THIS^.AddDataToContainer(ipData:=TurSt));
	W: FB_DO_WTURBINE_LD0_WTUR1_W := (sClass:='MV', bLinkResult:=THIS^.AddDataToContainer(ipData:=W));
	TurOp: FB_DO_WTURBINE_LD0_WTUR1_TurOp := (sClass:='CMD', bLinkResult:=THIS^.AddDataToContainer(ipData:=TurOp));
	DmdWSpt: FB_DO_WTURBINE_LD0_WTUR1_DmdWSpt := (sClass:='SPV', bLinkResult:=THIS^.AddDataToContainer(ipData:=DmdWSpt));
	TurCtl: FB_DO_WTURBINE_LD0_WTUR1_TurCtl := (sClass:='CMD', bLinkResult:=THIS^.AddDataToContainer(ipData:=TurCtl));
END_VAR
VAR
END_VAR

END_FUNCTION_BLOCK

